PROGRAM main
  VAR
    CONVEYOR_RUN AT %QX0.0 : BOOL;
    PUSHER_EXTEND AT %QX0.1 : BOOL;
    PUSHER_RETRACT AT %QX0.2 : BOOL;
    PASS_LAMP AT %QX0.3 : BOOL;
    FAIL_LAMP AT %QX0.4 : BOOL;
    FAULT_LAMP AT %QX0.5 : BOOL;
    STATION_READY AT %QX0.6 : BOOL;
    SIM_MODE AT %QX2.0 : BOOL := TRUE;
    SIM_UNIT_AT_INSPECTION AT %QX2.1 : BOOL := FALSE;
    SIM_UNIT_AT_REJECT AT %QX2.2 : BOOL := FALSE;
    SIM_VISION_PASS AT %QX2.3 : BOOL := FALSE;
    SIM_VISION_RESULT_VALID AT %QX2.4 : BOOL := FALSE;
    SIM_ESTOP_OK_NC AT %QX2.5 : BOOL := TRUE;
    SIM_GUARD_CLOSED_NC AT %QX2.6 : BOOL := TRUE;
    SIM_AUTO_MODE AT %QX2.7 : BOOL := TRUE;
    SIM_CYCLE_START AT %QX3.0 : BOOL := FALSE;
    SIM_RESET_PB AT %QX3.1 : BOOL := FALSE;
    SIM_PUSHER_EXTENDED AT %QX3.2 : BOOL := FALSE;
    SIM_PUSHER_RETRACTED AT %QX3.3 : BOOL := TRUE;
    SIM_DOWNSTREAM_CLEAR AT %QX3.4 : BOOL := TRUE;
    STATE_CODE AT %QW0 : UINT := 0;
    TOTAL_UNITS AT %QW1 : UINT := 0;
    TOTAL_REJECTS AT %QW2 : UINT := 0;
    LAST_CYCLE_TIME_MS AT %QW3 : UINT := 0;
    FAULT_CODE AT %QW4 : UINT := 0;
    LAST_SERIAL AT %QW5 : UINT := 0;
    LAST_RESULT AT %QW6 : UINT := 0;
    LAST_FAIL_REASON AT %QW7 : UINT := 0;
    SCENARIO_STEP AT %QW8 : UINT := 0;
    SIM_UNIT_SERIAL_IN AT %QW20 : UINT := 0;
    SIM_FAIL_REASON_IN AT %QW21 : UINT := 0;
    S_IDLE : BOOL := TRUE;
    S_READY : BOOL := FALSE;
    S_INSPECTING : BOOL := FALSE;
    S_PASS_RELEASE : BOOL := FALSE;
    S_REJECT_EXTEND : BOOL := FALSE;
    S_REJECT_RETRACT : BOOL := FALSE;
    S_FAULT : BOOL := FALSE;
    IN_UNIT_AT_INSPECTION : BOOL := FALSE;
    IN_UNIT_AT_REJECT : BOOL := FALSE;
    IN_VISION_PASS : BOOL := FALSE;
    IN_VISION_RESULT_VALID : BOOL := FALSE;
    IN_ESTOP_OK_NC : BOOL := FALSE;
    IN_GUARD_CLOSED_NC : BOOL := FALSE;
    IN_AUTO_MODE : BOOL := FALSE;
    IN_CYCLE_START : BOOL := FALSE;
    IN_RESET_PB : BOOL := FALSE;
    IN_PUSHER_EXTENDED : BOOL := FALSE;
    IN_PUSHER_RETRACTED : BOOL := FALSE;
    IN_DOWNSTREAM_CLEAR : BOOL := FALSE;
    START_RISE : BOOL := FALSE;
    START_LAST : BOOL := FALSE;
    RESET_RISE : BOOL := FALSE;
    RESET_LAST : BOOL := FALSE;
    UNIT_RISE : BOOL := FALSE;
    UNIT_LAST : BOOL := FALSE;
    VISION_LAST : BOOL := FALSE;
    VISION_CHANGED : BOOL := FALSE;
    VISION_UNSTABLE_LATCH : BOOL := FALSE;
    RESULT_LATCHED : BOOL := FALSE;
    RESULT_PASS_LATCH : BOOL := FALSE;
    RESULT_FAIL_LATCH : BOOL := FALSE;
    COMPLETE_PULSE : BOOL := FALSE;
    PASS_COMPLETE_PULSE : BOOL := FALSE;
    FAIL_COMPLETE_PULSE : BOOL := FALSE;
    EXTEND_DEMAND : BOOL := FALSE;
    RETRACT_DEMAND : BOOL := FALSE;
    OUTPUT_CONFLICT : BOOL := FALSE;
    FAULT_ESTOP : BOOL := FALSE;
    FAULT_GUARD : BOOL := FALSE;
    FAULT_EXTEND_TIMEOUT : BOOL := FALSE;
    FAULT_RETRACT_TIMEOUT : BOOL := FALSE;
    FAULT_UNIT_STUCK : BOOL := FALSE;
    FAULT_VISION_UNSTABLE : BOOL := FALSE;
    FAULT_OUTPUT_CONFLICT : BOOL := FALSE;
    UNIT_RELEASE_MONITOR : BOOL := FALSE;
    T_VISION_STABLE : TON;
    T_VISION_UNSTABLE : TON;
    T_PASS_RELEASE : TON;
    T_EXTEND_TIMEOUT : TON;
    T_REJECT_SETTLE : TON;
    T_RETRACT_TIMEOUT : TON;
    T_UNIT_STUCK : TON;
    IN_UNIT_SERIAL : UINT := 0;
    IN_FAIL_REASON : UINT := 0;
    CURRENT_SERIAL : UINT := 0;
    CURRENT_FAIL_REASON : UINT := 0;
    CYCLE_START_MS : UDINT := 0;
    NOW_MS : UDINT := 0;
    ALL_SAFE : BOOL := FALSE;
    TON0 : TON;
    TON1 : TON;
    TON2 : TON;
    TON3 : TON;
    TON4 : TON;
    TON5 : TON;
    TON6 : TON;
    TON7 : TON;
    TON8 : TON;
    TON9 : TON;
  END_VAR

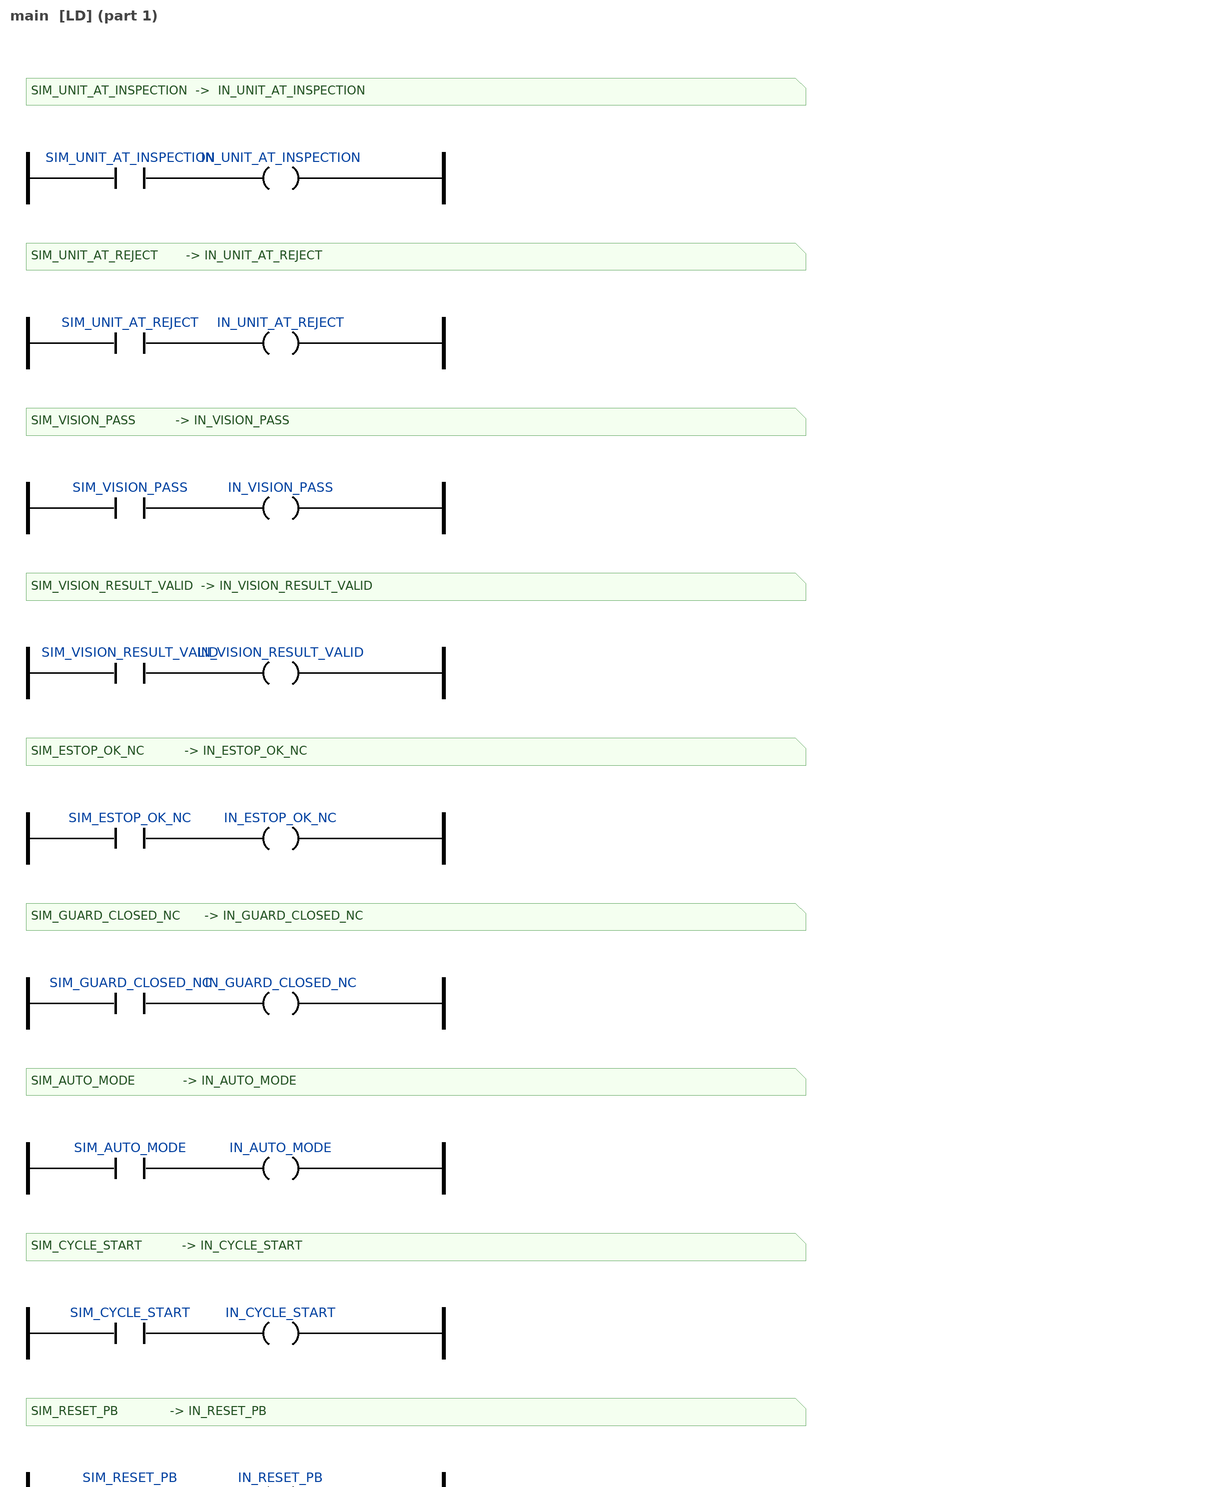
(* LD diagram, written out as Structured Text *)
(* SIM_UNIT_AT_INSPECTION  ->  IN_UNIT_AT_INSPECTION *)
IN_UNIT_AT_INSPECTION := SIM_UNIT_AT_INSPECTION;
(* SIM_UNIT_AT_REJECT       -> IN_UNIT_AT_REJECT *)
IN_UNIT_AT_REJECT := SIM_UNIT_AT_REJECT;
(* SIM_VISION_PASS          -> IN_VISION_PASS *)
IN_VISION_PASS := SIM_VISION_PASS;
(* SIM_VISION_RESULT_VALID  -> IN_VISION_RESULT_VALID *)
IN_VISION_RESULT_VALID := SIM_VISION_RESULT_VALID;
(* SIM_ESTOP_OK_NC          -> IN_ESTOP_OK_NC *)
IN_ESTOP_OK_NC := SIM_ESTOP_OK_NC;
(* SIM_GUARD_CLOSED_NC      -> IN_GUARD_CLOSED_NC *)
IN_GUARD_CLOSED_NC := SIM_GUARD_CLOSED_NC;
(* SIM_AUTO_MODE            -> IN_AUTO_MODE *)
IN_AUTO_MODE := SIM_AUTO_MODE;
(* SIM_CYCLE_START          -> IN_CYCLE_START *)
IN_CYCLE_START := SIM_CYCLE_START;
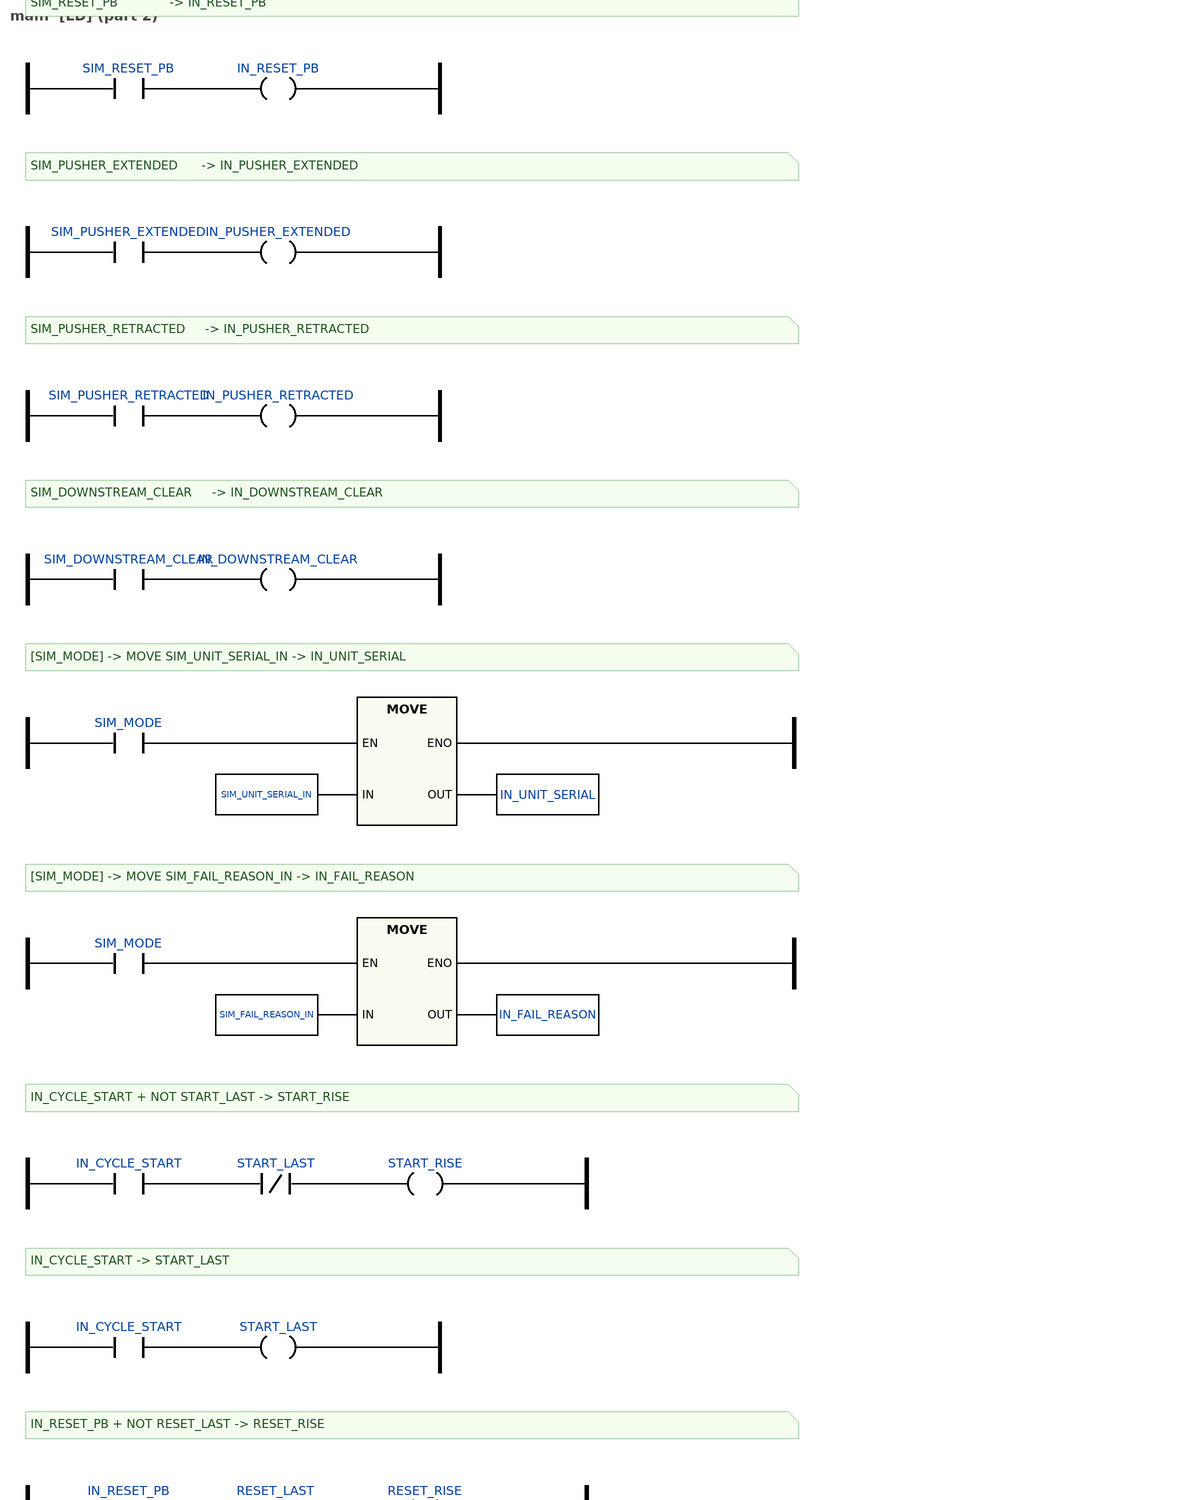
(* SIM_RESET_PB             -> IN_RESET_PB *)
IN_RESET_PB := SIM_RESET_PB;
(* SIM_PUSHER_EXTENDED      -> IN_PUSHER_EXTENDED *)
IN_PUSHER_EXTENDED := SIM_PUSHER_EXTENDED;
(* SIM_PUSHER_RETRACTED     -> IN_PUSHER_RETRACTED *)
IN_PUSHER_RETRACTED := SIM_PUSHER_RETRACTED;
(* SIM_DOWNSTREAM_CLEAR     -> IN_DOWNSTREAM_CLEAR *)
IN_DOWNSTREAM_CLEAR := SIM_DOWNSTREAM_CLEAR;
(* [SIM_MODE] -> MOVE SIM_UNIT_SERIAL_IN -> IN_UNIT_SERIAL *)
IF SIM_MODE THEN IN_UNIT_SERIAL := SIM_UNIT_SERIAL_IN; END_IF;
(* [SIM_MODE] -> MOVE SIM_FAIL_REASON_IN -> IN_FAIL_REASON *)
IF SIM_MODE THEN IN_FAIL_REASON := SIM_FAIL_REASON_IN; END_IF;
(* IN_CYCLE_START + NOT START_LAST -> START_RISE *)
START_RISE := IN_CYCLE_START AND NOT START_LAST;
(* IN_CYCLE_START -> START_LAST *)
START_LAST := IN_CYCLE_START;
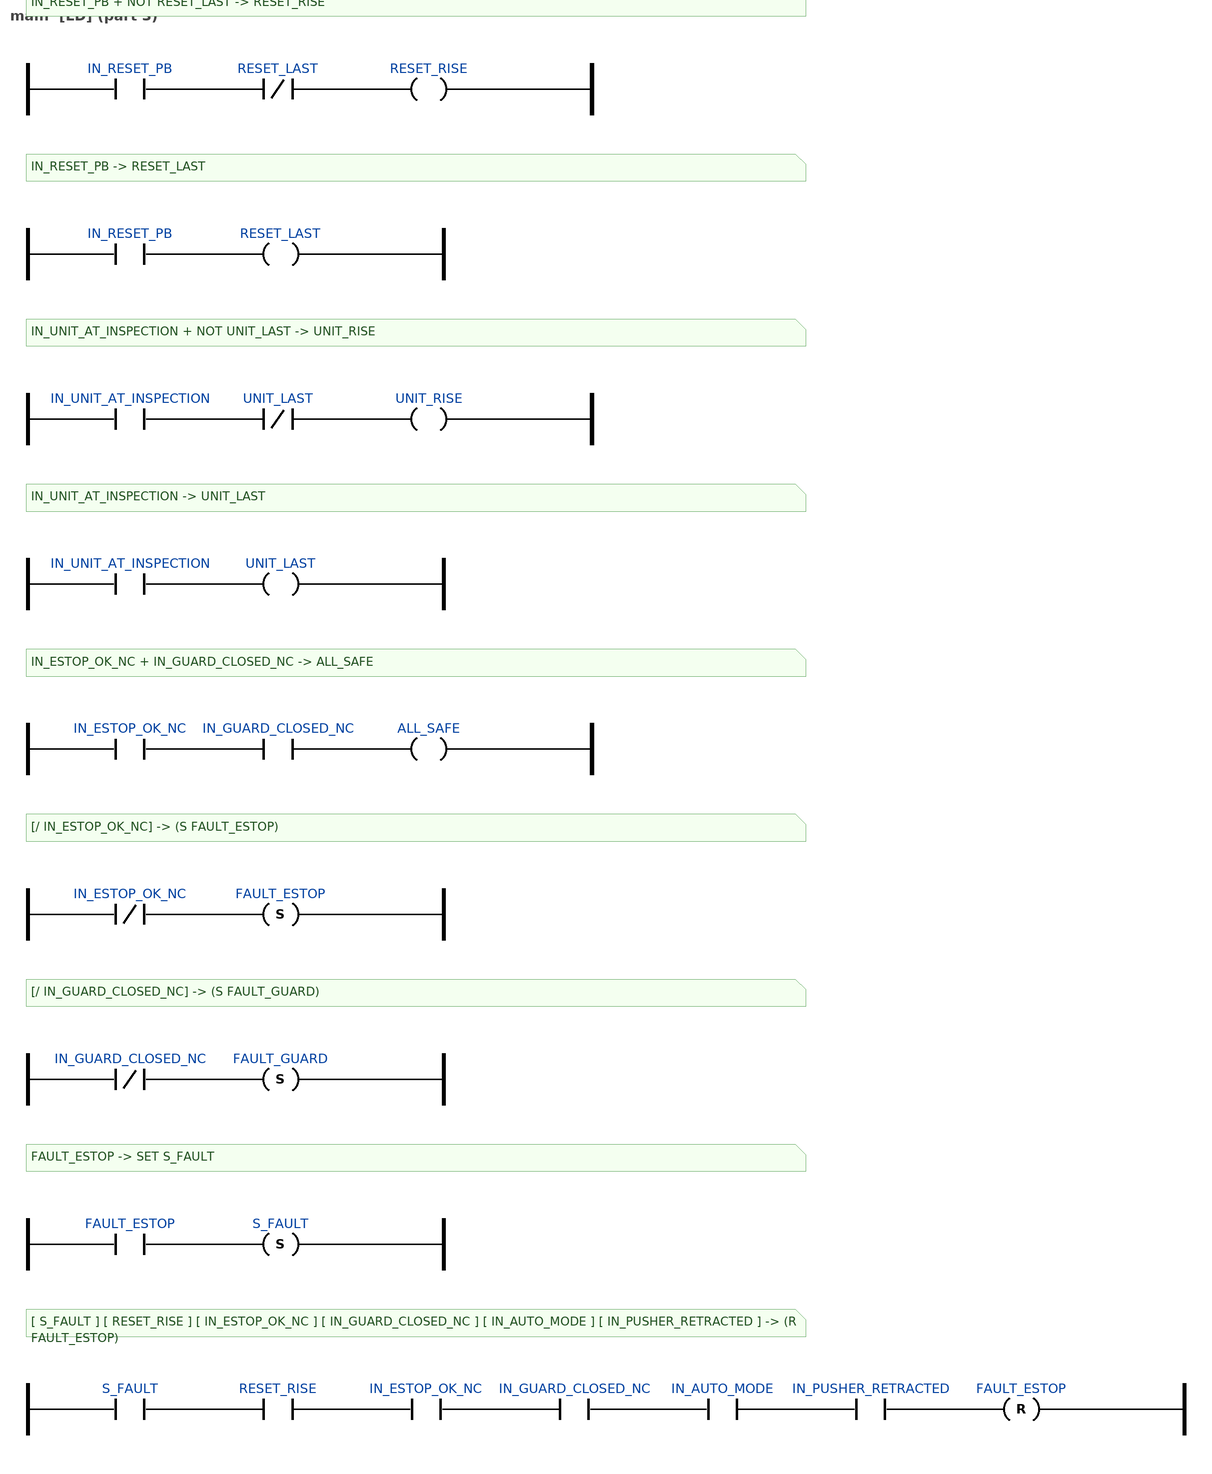
(* IN_RESET_PB + NOT RESET_LAST -> RESET_RISE *)
RESET_RISE := IN_RESET_PB AND NOT RESET_LAST;
(* IN_RESET_PB -> RESET_LAST *)
RESET_LAST := IN_RESET_PB;
(* IN_UNIT_AT_INSPECTION + NOT UNIT_LAST -> UNIT_RISE *)
UNIT_RISE := IN_UNIT_AT_INSPECTION AND NOT UNIT_LAST;
(* IN_UNIT_AT_INSPECTION -> UNIT_LAST *)
UNIT_LAST := IN_UNIT_AT_INSPECTION;
(* IN_ESTOP_OK_NC + IN_GUARD_CLOSED_NC -> ALL_SAFE *)
ALL_SAFE := IN_ESTOP_OK_NC AND IN_GUARD_CLOSED_NC;
(* [/ IN_ESTOP_OK_NC] -> (S FAULT_ESTOP) *)
IF NOT IN_ESTOP_OK_NC THEN FAULT_ESTOP := TRUE; END_IF;
(* [/ IN_GUARD_CLOSED_NC] -> (S FAULT_GUARD) *)
IF NOT IN_GUARD_CLOSED_NC THEN FAULT_GUARD := TRUE; END_IF;
(* FAULT_ESTOP -> SET S_FAULT *)
IF FAULT_ESTOP THEN S_FAULT := TRUE; END_IF;
(* [ S_FAULT ] [ RESET_RISE ] [ IN_ESTOP_OK_NC ] [ IN_GUARD_CLOSED_NC ] [ IN_AUTO_MODE ] [ IN_PUSHER_RETRACTED ] -> (R FAULT_ESTOP) *)
IF S_FAULT AND RESET_RISE AND IN_ESTOP_OK_NC AND IN_GUARD_CLOSED_NC AND IN_AUTO_MODE AND IN_PUSHER_RETRACTED THEN FAULT_ESTOP := FALSE; END_IF;
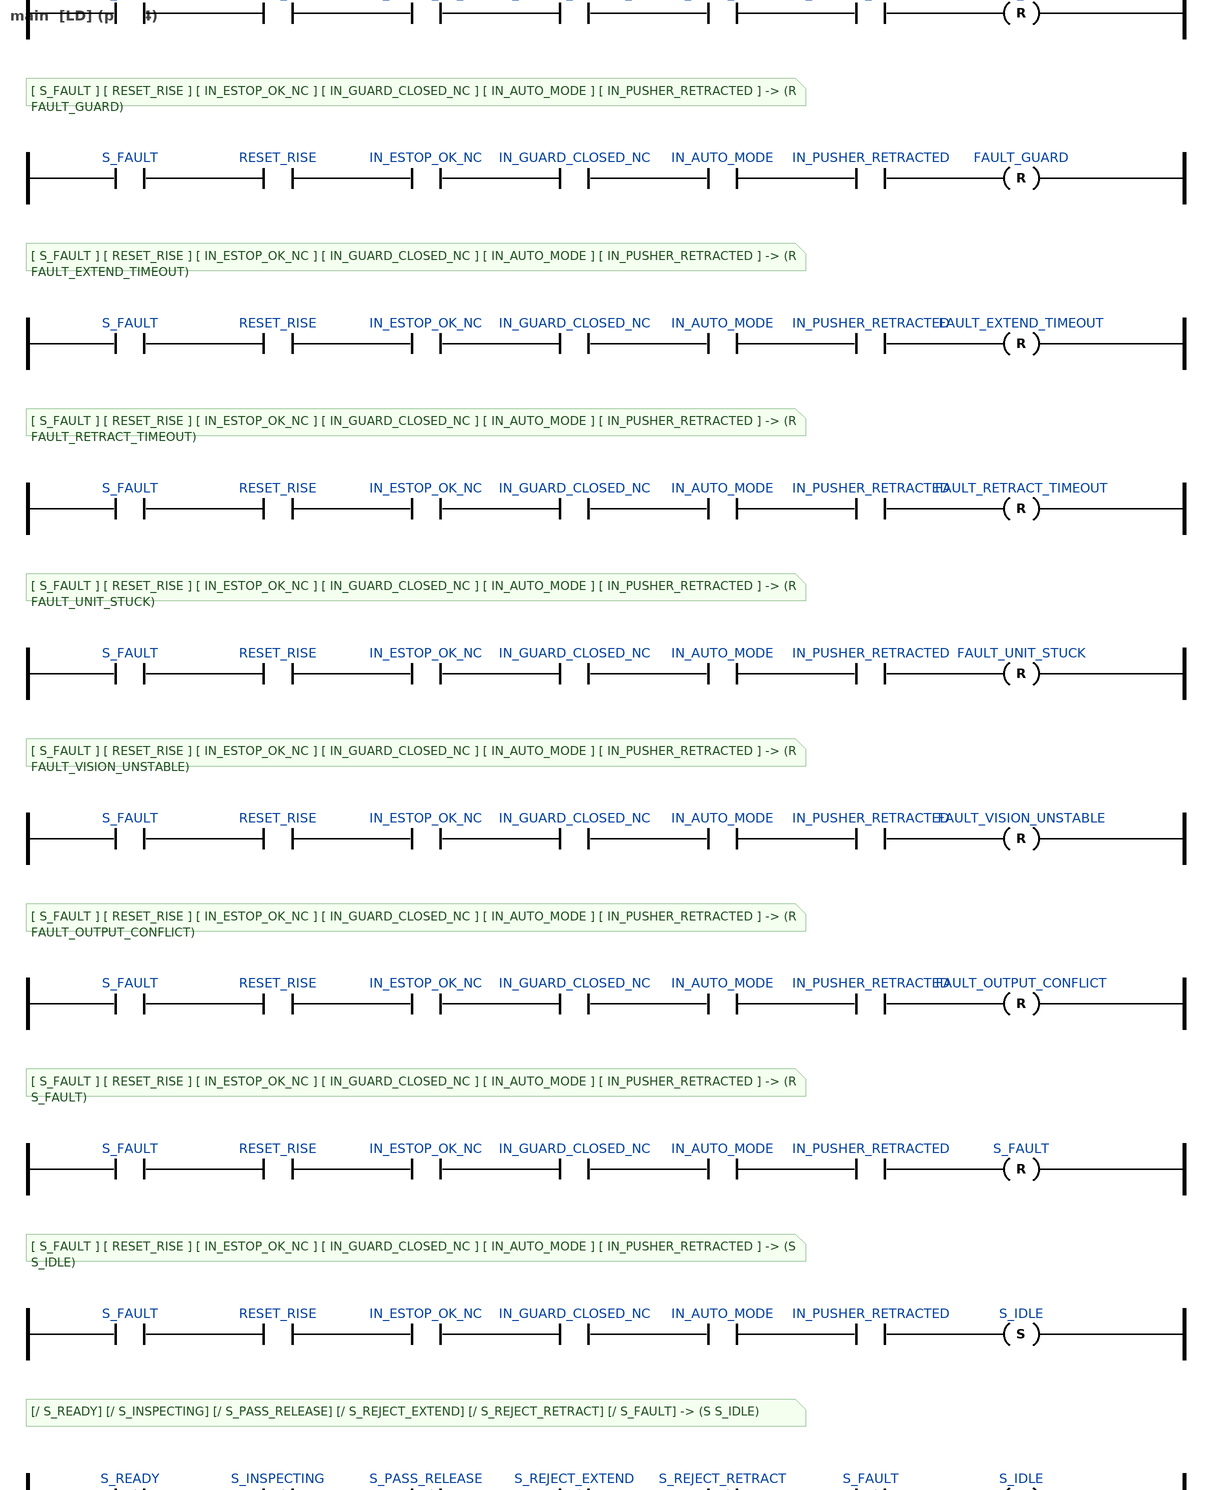
(* [ S_FAULT ] [ RESET_RISE ] [ IN_ESTOP_OK_NC ] [ IN_GUARD_CLOSED_NC ] [ IN_AUTO_MODE ] [ IN_PUSHER_RETRACTED ] -> (R FAULT_GUARD) *)
IF S_FAULT AND RESET_RISE AND IN_ESTOP_OK_NC AND IN_GUARD_CLOSED_NC AND IN_AUTO_MODE AND IN_PUSHER_RETRACTED THEN FAULT_GUARD := FALSE; END_IF;
(* [ S_FAULT ] [ RESET_RISE ] [ IN_ESTOP_OK_NC ] [ IN_GUARD_CLOSED_NC ] [ IN_AUTO_MODE ] [ IN_PUSHER_RETRACTED ] -> (R FAULT_EXTEND_TIMEOUT) *)
IF S_FAULT AND RESET_RISE AND IN_ESTOP_OK_NC AND IN_GUARD_CLOSED_NC AND IN_AUTO_MODE AND IN_PUSHER_RETRACTED THEN FAULT_EXTEND_TIMEOUT := FALSE; END_IF;
(* [ S_FAULT ] [ RESET_RISE ] [ IN_ESTOP_OK_NC ] [ IN_GUARD_CLOSED_NC ] [ IN_AUTO_MODE ] [ IN_PUSHER_RETRACTED ] -> (R FAULT_RETRACT_TIMEOUT) *)
IF S_FAULT AND RESET_RISE AND IN_ESTOP_OK_NC AND IN_GUARD_CLOSED_NC AND IN_AUTO_MODE AND IN_PUSHER_RETRACTED THEN FAULT_RETRACT_TIMEOUT := FALSE; END_IF;
(* [ S_FAULT ] [ RESET_RISE ] [ IN_ESTOP_OK_NC ] [ IN_GUARD_CLOSED_NC ] [ IN_AUTO_MODE ] [ IN_PUSHER_RETRACTED ] -> (R FAULT_UNIT_STUCK) *)
IF S_FAULT AND RESET_RISE AND IN_ESTOP_OK_NC AND IN_GUARD_CLOSED_NC AND IN_AUTO_MODE AND IN_PUSHER_RETRACTED THEN FAULT_UNIT_STUCK := FALSE; END_IF;
(* [ S_FAULT ] [ RESET_RISE ] [ IN_ESTOP_OK_NC ] [ IN_GUARD_CLOSED_NC ] [ IN_AUTO_MODE ] [ IN_PUSHER_RETRACTED ] -> (R FAULT_VISION_UNSTABLE) *)
IF S_FAULT AND RESET_RISE AND IN_ESTOP_OK_NC AND IN_GUARD_CLOSED_NC AND IN_AUTO_MODE AND IN_PUSHER_RETRACTED THEN FAULT_VISION_UNSTABLE := FALSE; END_IF;
(* [ S_FAULT ] [ RESET_RISE ] [ IN_ESTOP_OK_NC ] [ IN_GUARD_CLOSED_NC ] [ IN_AUTO_MODE ] [ IN_PUSHER_RETRACTED ] -> (R FAULT_OUTPUT_CONFLICT) *)
IF S_FAULT AND RESET_RISE AND IN_ESTOP_OK_NC AND IN_GUARD_CLOSED_NC AND IN_AUTO_MODE AND IN_PUSHER_RETRACTED THEN FAULT_OUTPUT_CONFLICT := FALSE; END_IF;
(* [ S_FAULT ] [ RESET_RISE ] [ IN_ESTOP_OK_NC ] [ IN_GUARD_CLOSED_NC ] [ IN_AUTO_MODE ] [ IN_PUSHER_RETRACTED ] -> (R S_FAULT) *)
IF S_FAULT AND RESET_RISE AND IN_ESTOP_OK_NC AND IN_GUARD_CLOSED_NC AND IN_AUTO_MODE AND IN_PUSHER_RETRACTED THEN S_FAULT := FALSE; END_IF;
(* [ S_FAULT ] [ RESET_RISE ] [ IN_ESTOP_OK_NC ] [ IN_GUARD_CLOSED_NC ] [ IN_AUTO_MODE ] [ IN_PUSHER_RETRACTED ] -> (S S_IDLE) *)
IF S_FAULT AND RESET_RISE AND IN_ESTOP_OK_NC AND IN_GUARD_CLOSED_NC AND IN_AUTO_MODE AND IN_PUSHER_RETRACTED THEN S_IDLE := TRUE; END_IF;
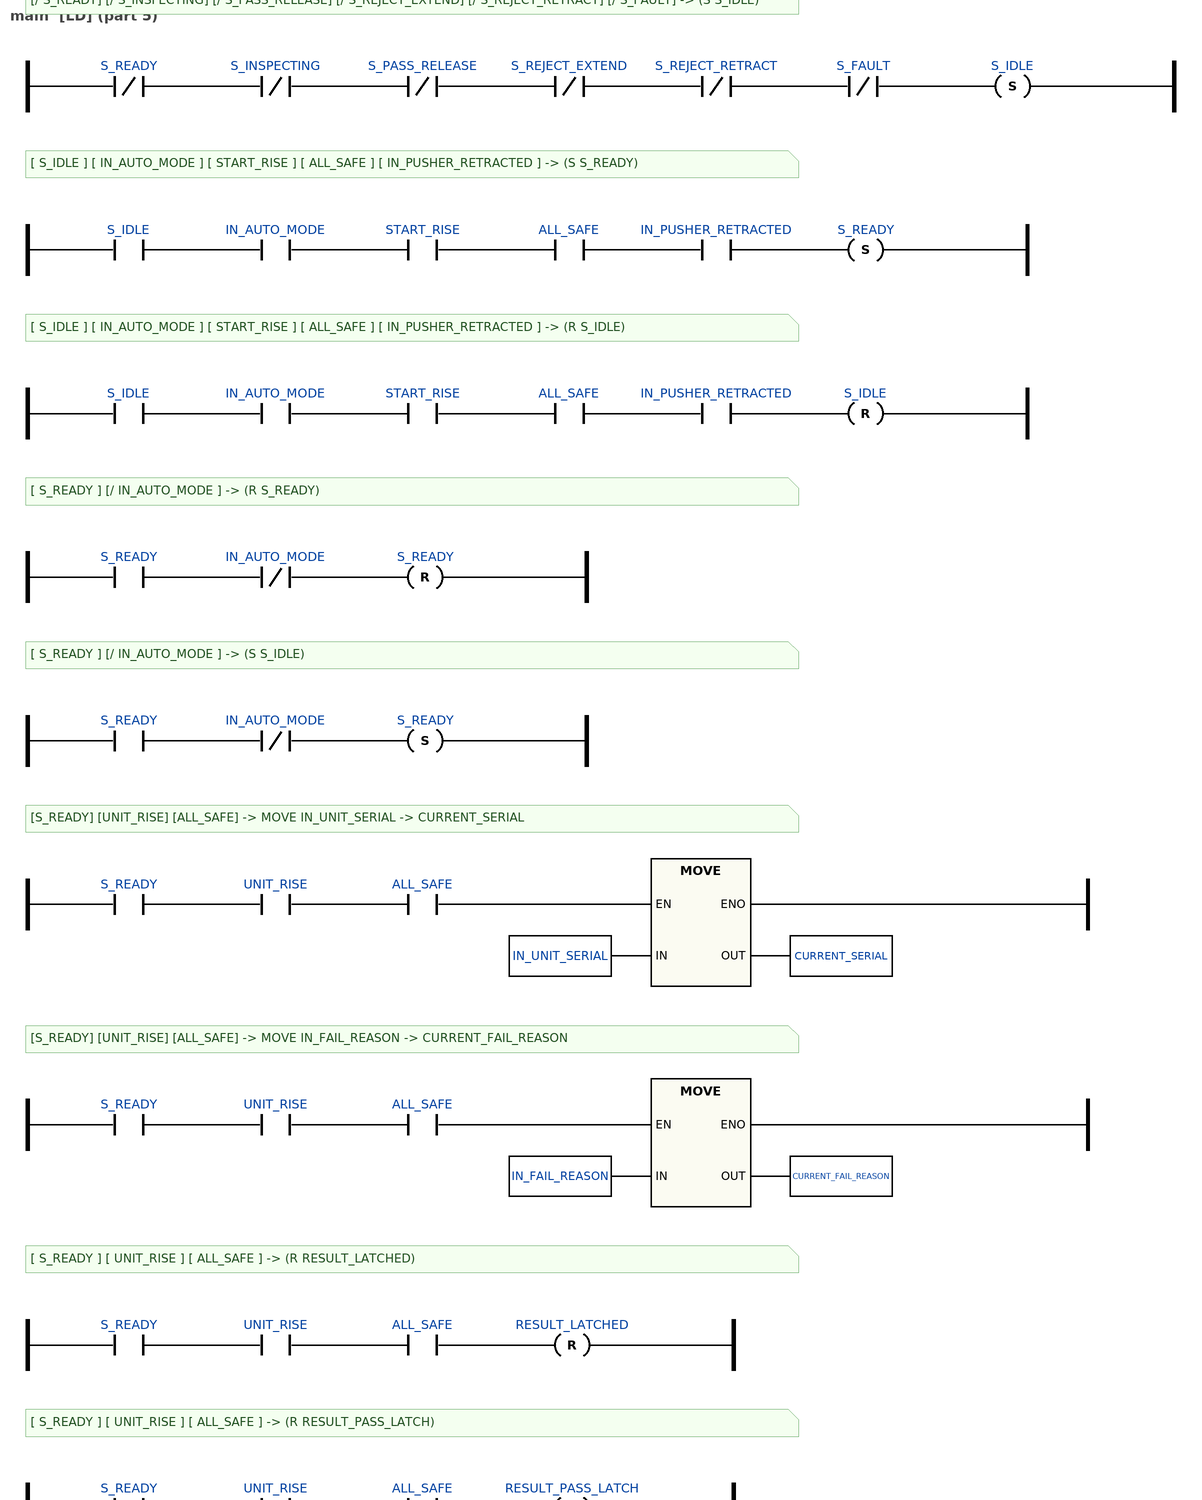
(* [/ S_READY] [/ S_INSPECTING] [/ S_PASS_RELEASE] [/ S_REJECT_EXTEND] [/ S_REJECT_RETRACT] [/ S_FAULT] -> (S S_IDLE) *)
IF NOT S_READY AND NOT S_INSPECTING AND NOT S_PASS_RELEASE AND NOT S_REJECT_EXTEND AND NOT S_REJECT_RETRACT AND NOT S_FAULT THEN S_IDLE := TRUE; END_IF;
(* [ S_IDLE ] [ IN_AUTO_MODE ] [ START_RISE ] [ ALL_SAFE ] [ IN_PUSHER_RETRACTED ] -> (S S_READY) *)
IF S_IDLE AND IN_AUTO_MODE AND START_RISE AND ALL_SAFE AND IN_PUSHER_RETRACTED THEN S_READY := TRUE; END_IF;
(* [ S_IDLE ] [ IN_AUTO_MODE ] [ START_RISE ] [ ALL_SAFE ] [ IN_PUSHER_RETRACTED ] -> (R S_IDLE) *)
IF S_IDLE AND IN_AUTO_MODE AND START_RISE AND ALL_SAFE AND IN_PUSHER_RETRACTED THEN S_IDLE := FALSE; END_IF;
(* [ S_READY ] [/ IN_AUTO_MODE ] -> (R S_READY) *)
IF S_READY AND NOT IN_AUTO_MODE THEN S_READY := FALSE; END_IF;
(* [ S_READY ] [/ IN_AUTO_MODE ] -> (S S_IDLE) *)
IF S_READY AND NOT IN_AUTO_MODE THEN S_READY := TRUE; END_IF;
(* [S_READY] [UNIT_RISE] [ALL_SAFE] -> MOVE IN_UNIT_SERIAL -> CURRENT_SERIAL *)
IF S_READY AND UNIT_RISE AND ALL_SAFE THEN CURRENT_SERIAL := IN_UNIT_SERIAL; END_IF;
(* [S_READY] [UNIT_RISE] [ALL_SAFE] -> MOVE IN_FAIL_REASON -> CURRENT_FAIL_REASON *)
IF S_READY AND UNIT_RISE AND ALL_SAFE THEN CURRENT_FAIL_REASON := IN_FAIL_REASON; END_IF;
(* [ S_READY ] [ UNIT_RISE ] [ ALL_SAFE ] -> (R RESULT_LATCHED) *)
IF S_READY AND UNIT_RISE AND ALL_SAFE THEN RESULT_LATCHED := FALSE; END_IF;
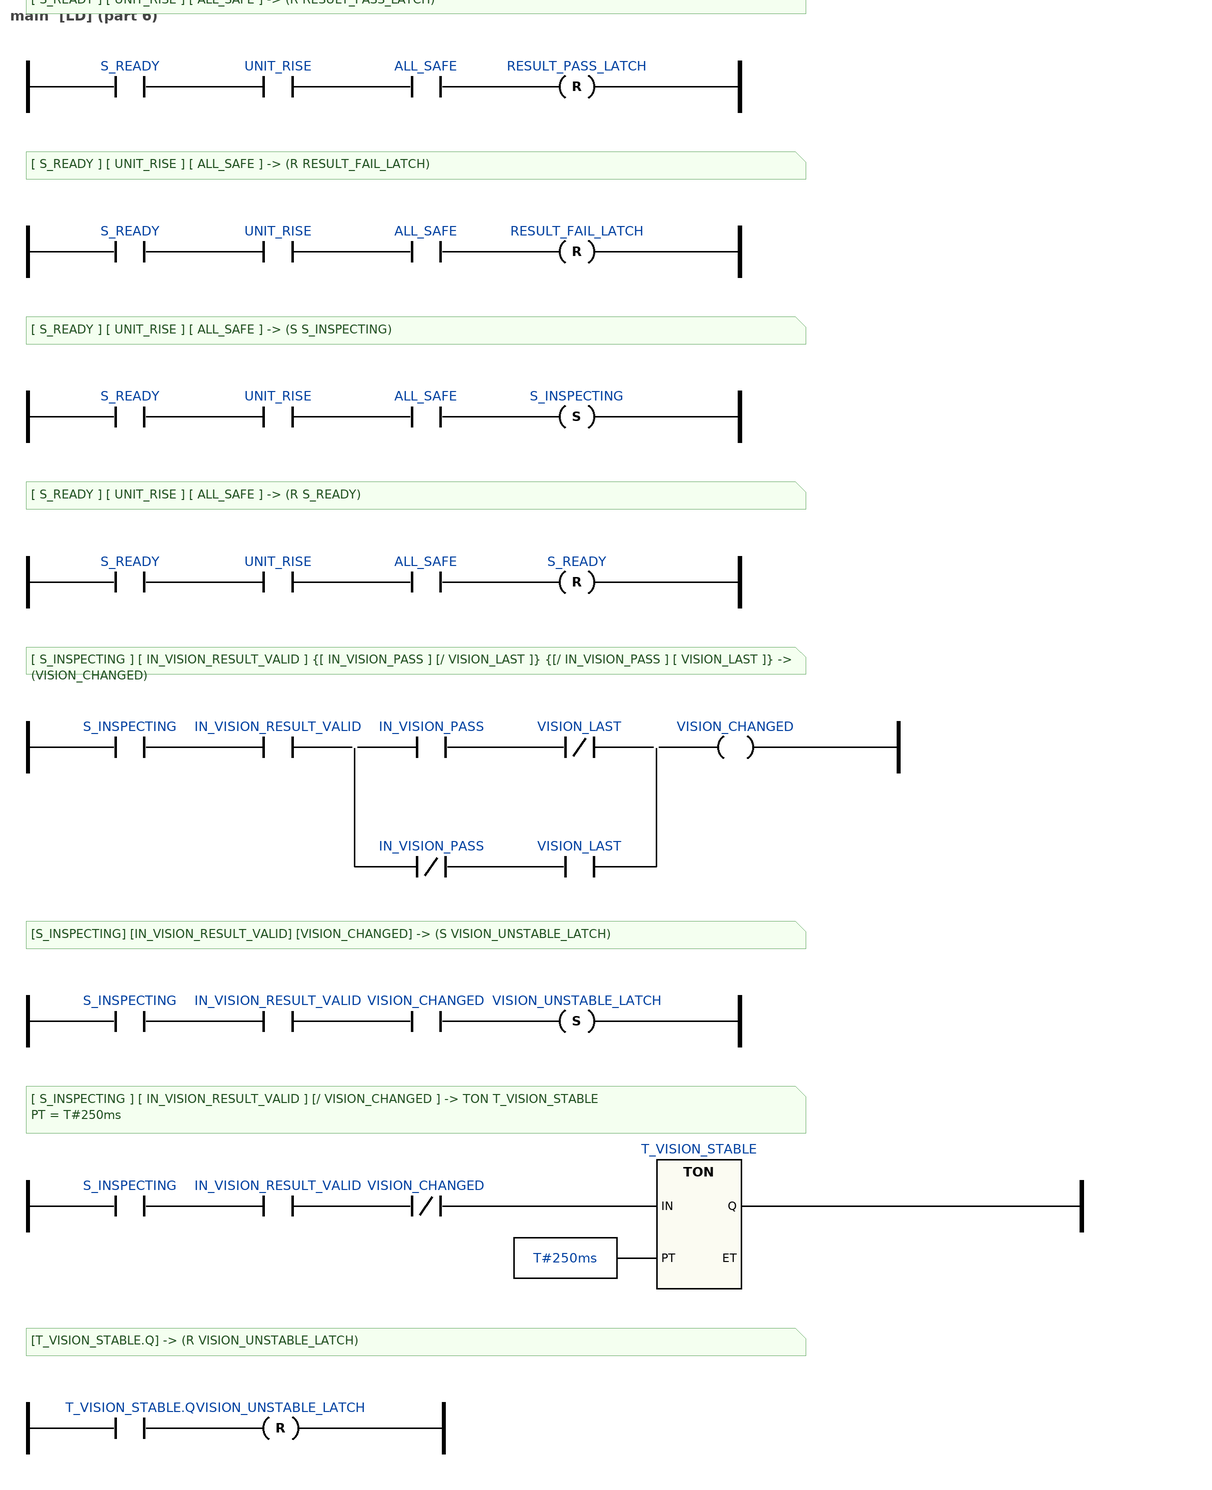
(* [ S_READY ] [ UNIT_RISE ] [ ALL_SAFE ] -> (R RESULT_PASS_LATCH) *)
IF S_READY AND UNIT_RISE AND ALL_SAFE THEN RESULT_PASS_LATCH := FALSE; END_IF;
(* [ S_READY ] [ UNIT_RISE ] [ ALL_SAFE ] -> (R RESULT_FAIL_LATCH) *)
IF S_READY AND UNIT_RISE AND ALL_SAFE THEN RESULT_FAIL_LATCH := FALSE; END_IF;
(* [ S_READY ] [ UNIT_RISE ] [ ALL_SAFE ] -> (S S_INSPECTING) *)
IF S_READY AND UNIT_RISE AND ALL_SAFE THEN S_INSPECTING := TRUE; END_IF;
(* [ S_READY ] [ UNIT_RISE ] [ ALL_SAFE ] -> (R S_READY) *)
IF S_READY AND UNIT_RISE AND ALL_SAFE THEN S_READY := FALSE; END_IF;
(* [ S_INSPECTING ] [ IN_VISION_RESULT_VALID ] {[ IN_VISION_PASS ] [/ VISION_LAST ]} {[/ IN_VISION_PASS ] [ VISION_LAST ]} -> (VISION_CHANGED) *)
VISION_CHANGED := S_INSPECTING AND IN_VISION_RESULT_VALID AND (NOT IN_VISION_PASS AND VISION_LAST OR IN_VISION_PASS AND NOT VISION_LAST);
(* [S_INSPECTING] [IN_VISION_RESULT_VALID] [VISION_CHANGED] -> (S VISION_UNSTABLE_LATCH) *)
IF S_INSPECTING AND IN_VISION_RESULT_VALID AND VISION_CHANGED THEN VISION_UNSTABLE_LATCH := TRUE; END_IF;
(* [ S_INSPECTING ] [ IN_VISION_RESULT_VALID ] [/ VISION_CHANGED ] -> TON T_VISION_STABLE
PT = T#250ms *)
(* [T_VISION_STABLE.Q] -> (R VISION_UNSTABLE_LATCH) *)
IF T_VISION_STABLE.Q THEN VISION_UNSTABLE_LATCH := FALSE; END_IF;
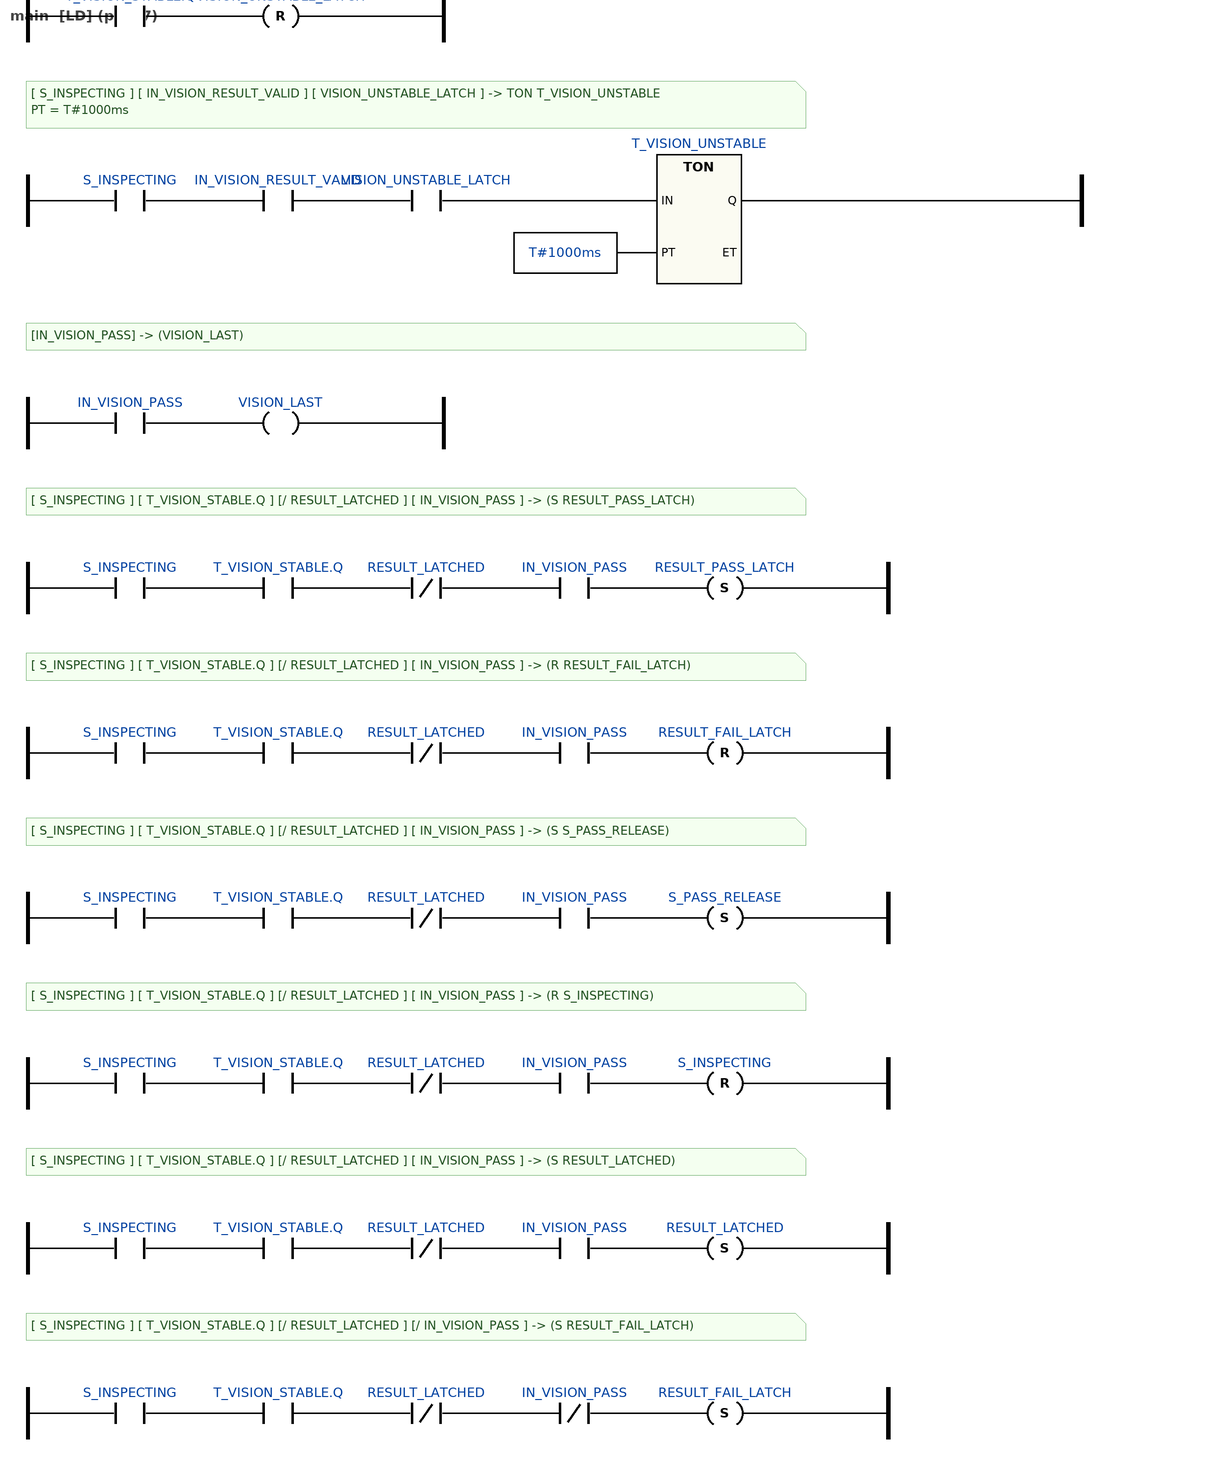
(* [ S_INSPECTING ] [ IN_VISION_RESULT_VALID ] [ VISION_UNSTABLE_LATCH ] -> TON T_VISION_UNSTABLE
PT = T#1000ms *)
(* [IN_VISION_PASS] -> (VISION_LAST) *)
VISION_LAST := IN_VISION_PASS;
(* [ S_INSPECTING ] [ T_VISION_STABLE.Q ] [/ RESULT_LATCHED ] [ IN_VISION_PASS ] -> (S RESULT_PASS_LATCH) *)
IF S_INSPECTING AND T_VISION_STABLE.Q AND NOT RESULT_LATCHED AND IN_VISION_PASS THEN RESULT_PASS_LATCH := TRUE; END_IF;
(* [ S_INSPECTING ] [ T_VISION_STABLE.Q ] [/ RESULT_LATCHED ] [ IN_VISION_PASS ] -> (R RESULT_FAIL_LATCH) *)
IF S_INSPECTING AND T_VISION_STABLE.Q AND NOT RESULT_LATCHED AND IN_VISION_PASS THEN RESULT_FAIL_LATCH := FALSE; END_IF;
(* [ S_INSPECTING ] [ T_VISION_STABLE.Q ] [/ RESULT_LATCHED ] [ IN_VISION_PASS ] -> (S S_PASS_RELEASE) *)
IF S_INSPECTING AND T_VISION_STABLE.Q AND NOT RESULT_LATCHED AND IN_VISION_PASS THEN S_PASS_RELEASE := TRUE; END_IF;
(* [ S_INSPECTING ] [ T_VISION_STABLE.Q ] [/ RESULT_LATCHED ] [ IN_VISION_PASS ] -> (R S_INSPECTING) *)
IF S_INSPECTING AND T_VISION_STABLE.Q AND NOT RESULT_LATCHED AND IN_VISION_PASS THEN S_INSPECTING := FALSE; END_IF;
(* [ S_INSPECTING ] [ T_VISION_STABLE.Q ] [/ RESULT_LATCHED ] [ IN_VISION_PASS ] -> (S RESULT_LATCHED) *)
IF S_INSPECTING AND T_VISION_STABLE.Q AND NOT RESULT_LATCHED AND IN_VISION_PASS THEN RESULT_LATCHED := TRUE; END_IF;
(* [ S_INSPECTING ] [ T_VISION_STABLE.Q ] [/ RESULT_LATCHED ] [/ IN_VISION_PASS ] -> (S RESULT_FAIL_LATCH) *)
IF S_INSPECTING AND T_VISION_STABLE.Q AND NOT RESULT_LATCHED AND NOT IN_VISION_PASS THEN RESULT_FAIL_LATCH := TRUE; END_IF;
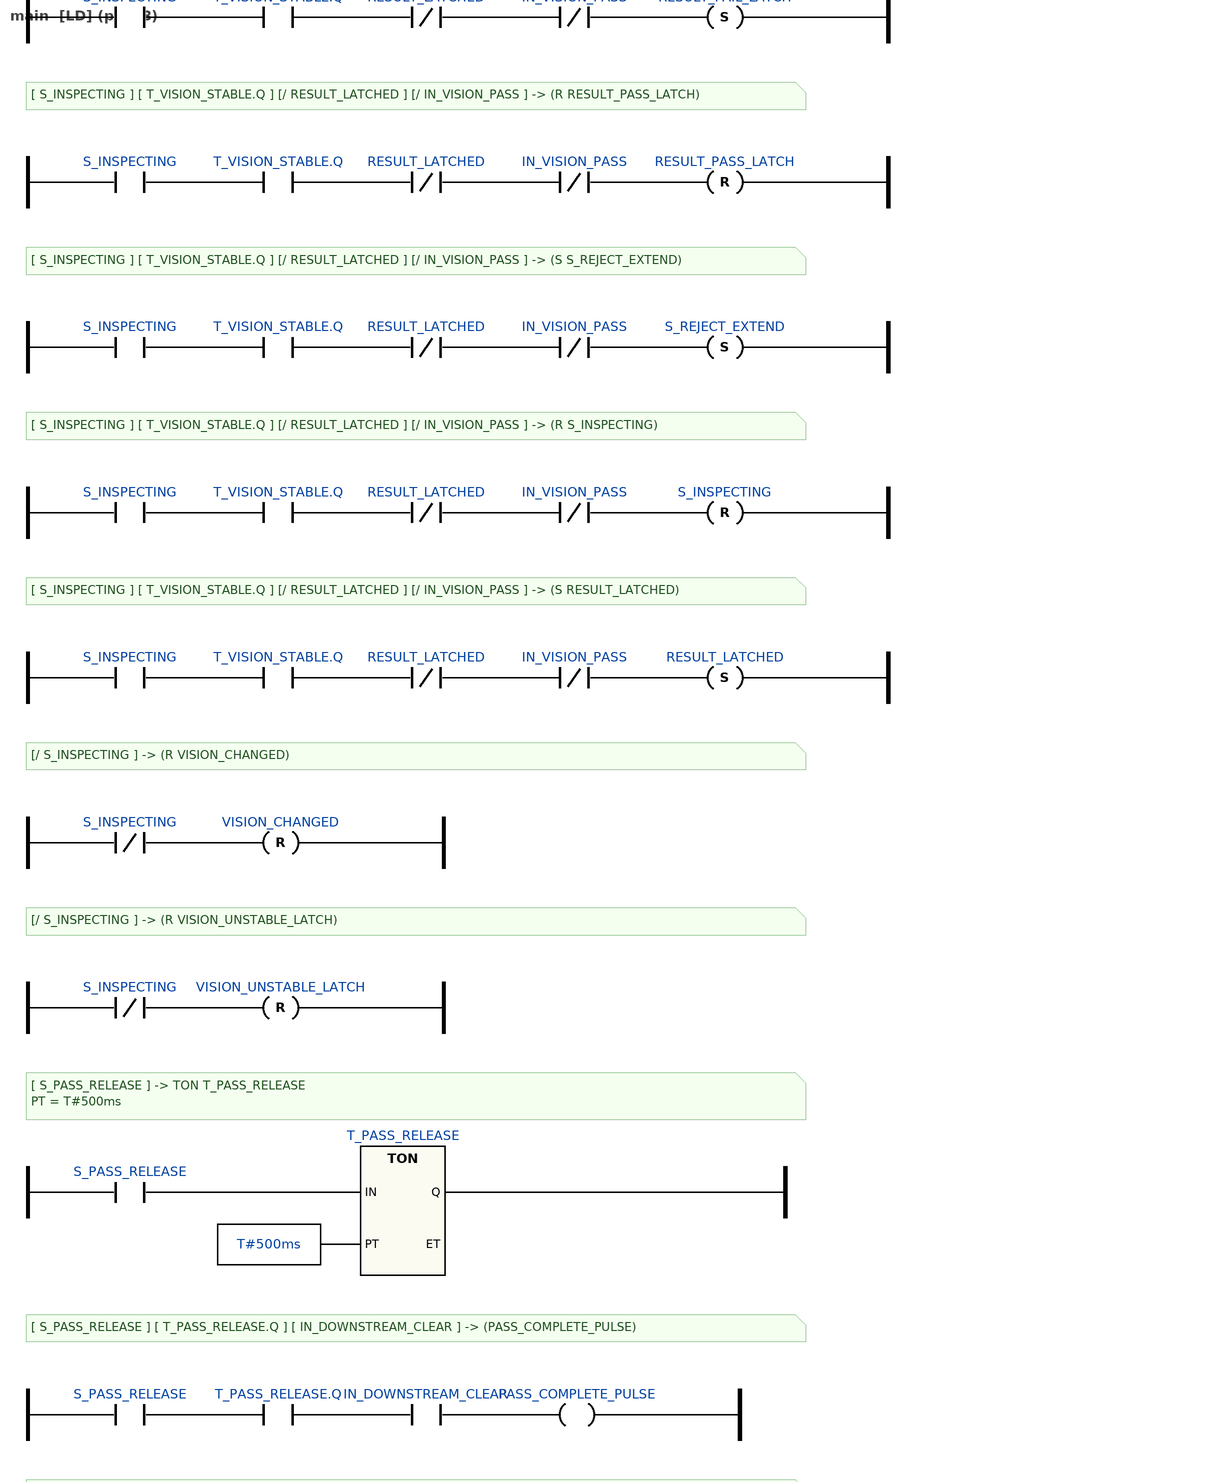
(* [ S_INSPECTING ] [ T_VISION_STABLE.Q ] [/ RESULT_LATCHED ] [/ IN_VISION_PASS ] -> (R RESULT_PASS_LATCH) *)
IF S_INSPECTING AND T_VISION_STABLE.Q AND NOT RESULT_LATCHED AND NOT IN_VISION_PASS THEN RESULT_PASS_LATCH := FALSE; END_IF;
(* [ S_INSPECTING ] [ T_VISION_STABLE.Q ] [/ RESULT_LATCHED ] [/ IN_VISION_PASS ] -> (S S_REJECT_EXTEND) *)
IF S_INSPECTING AND T_VISION_STABLE.Q AND NOT RESULT_LATCHED AND NOT IN_VISION_PASS THEN S_REJECT_EXTEND := TRUE; END_IF;
(* [ S_INSPECTING ] [ T_VISION_STABLE.Q ] [/ RESULT_LATCHED ] [/ IN_VISION_PASS ] -> (R S_INSPECTING) *)
IF S_INSPECTING AND T_VISION_STABLE.Q AND NOT RESULT_LATCHED AND NOT IN_VISION_PASS THEN S_INSPECTING := FALSE; END_IF;
(* [ S_INSPECTING ] [ T_VISION_STABLE.Q ] [/ RESULT_LATCHED ] [/ IN_VISION_PASS ] -> (S RESULT_LATCHED) *)
IF S_INSPECTING AND T_VISION_STABLE.Q AND NOT RESULT_LATCHED AND NOT IN_VISION_PASS THEN RESULT_LATCHED := TRUE; END_IF;
(* [/ S_INSPECTING ] -> (R VISION_CHANGED) *)
IF NOT S_INSPECTING THEN VISION_CHANGED := FALSE; END_IF;
(* [/ S_INSPECTING ] -> (R VISION_UNSTABLE_LATCH) *)
IF NOT S_INSPECTING THEN VISION_UNSTABLE_LATCH := FALSE; END_IF;
(* [ S_PASS_RELEASE ] -> TON T_PASS_RELEASE
PT = T#500ms *)
(* [ S_PASS_RELEASE ] [ T_PASS_RELEASE.Q ] [ IN_DOWNSTREAM_CLEAR ] -> (PASS_COMPLETE_PULSE) *)
PASS_COMPLETE_PULSE := S_PASS_RELEASE AND T_PASS_RELEASE.Q AND IN_DOWNSTREAM_CLEAR;
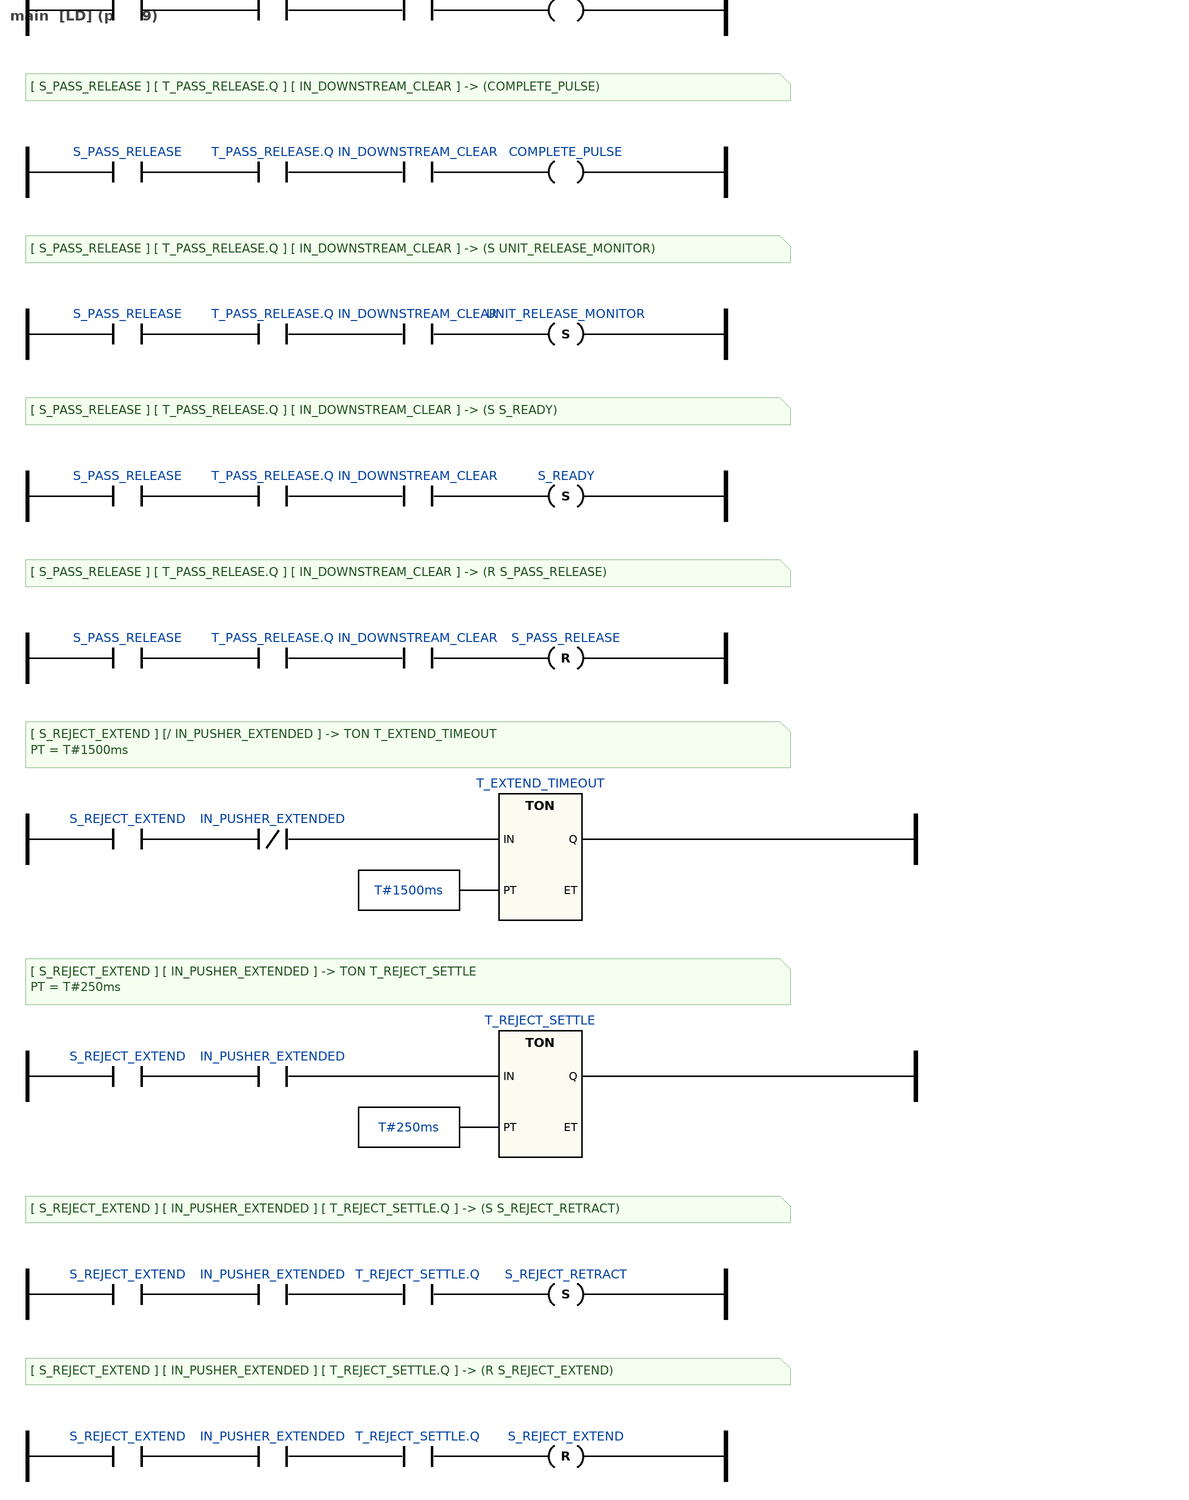
(* [ S_PASS_RELEASE ] [ T_PASS_RELEASE.Q ] [ IN_DOWNSTREAM_CLEAR ] -> (COMPLETE_PULSE) *)
COMPLETE_PULSE := S_PASS_RELEASE AND T_PASS_RELEASE.Q AND IN_DOWNSTREAM_CLEAR;
(* [ S_PASS_RELEASE ] [ T_PASS_RELEASE.Q ] [ IN_DOWNSTREAM_CLEAR ] -> (S UNIT_RELEASE_MONITOR) *)
IF S_PASS_RELEASE AND T_PASS_RELEASE.Q AND IN_DOWNSTREAM_CLEAR THEN UNIT_RELEASE_MONITOR := TRUE; END_IF;
(* [ S_PASS_RELEASE ] [ T_PASS_RELEASE.Q ] [ IN_DOWNSTREAM_CLEAR ] -> (S S_READY) *)
IF S_PASS_RELEASE AND T_PASS_RELEASE.Q AND IN_DOWNSTREAM_CLEAR THEN S_READY := TRUE; END_IF;
(* [ S_PASS_RELEASE ] [ T_PASS_RELEASE.Q ] [ IN_DOWNSTREAM_CLEAR ] -> (R S_PASS_RELEASE) *)
IF S_PASS_RELEASE AND T_PASS_RELEASE.Q AND IN_DOWNSTREAM_CLEAR THEN S_PASS_RELEASE := FALSE; END_IF;
(* [ S_REJECT_EXTEND ] [/ IN_PUSHER_EXTENDED ] -> TON T_EXTEND_TIMEOUT
PT = T#1500ms *)
(* [ S_REJECT_EXTEND ] [ IN_PUSHER_EXTENDED ] -> TON T_REJECT_SETTLE
PT = T#250ms *)
(* [ S_REJECT_EXTEND ] [ IN_PUSHER_EXTENDED ] [ T_REJECT_SETTLE.Q ] -> (S S_REJECT_RETRACT) *)
IF S_REJECT_EXTEND AND IN_PUSHER_EXTENDED AND T_REJECT_SETTLE.Q THEN S_REJECT_RETRACT := TRUE; END_IF;
(* [ S_REJECT_EXTEND ] [ IN_PUSHER_EXTENDED ] [ T_REJECT_SETTLE.Q ] -> (R S_REJECT_EXTEND) *)
IF S_REJECT_EXTEND AND IN_PUSHER_EXTENDED AND T_REJECT_SETTLE.Q THEN S_REJECT_EXTEND := FALSE; END_IF;
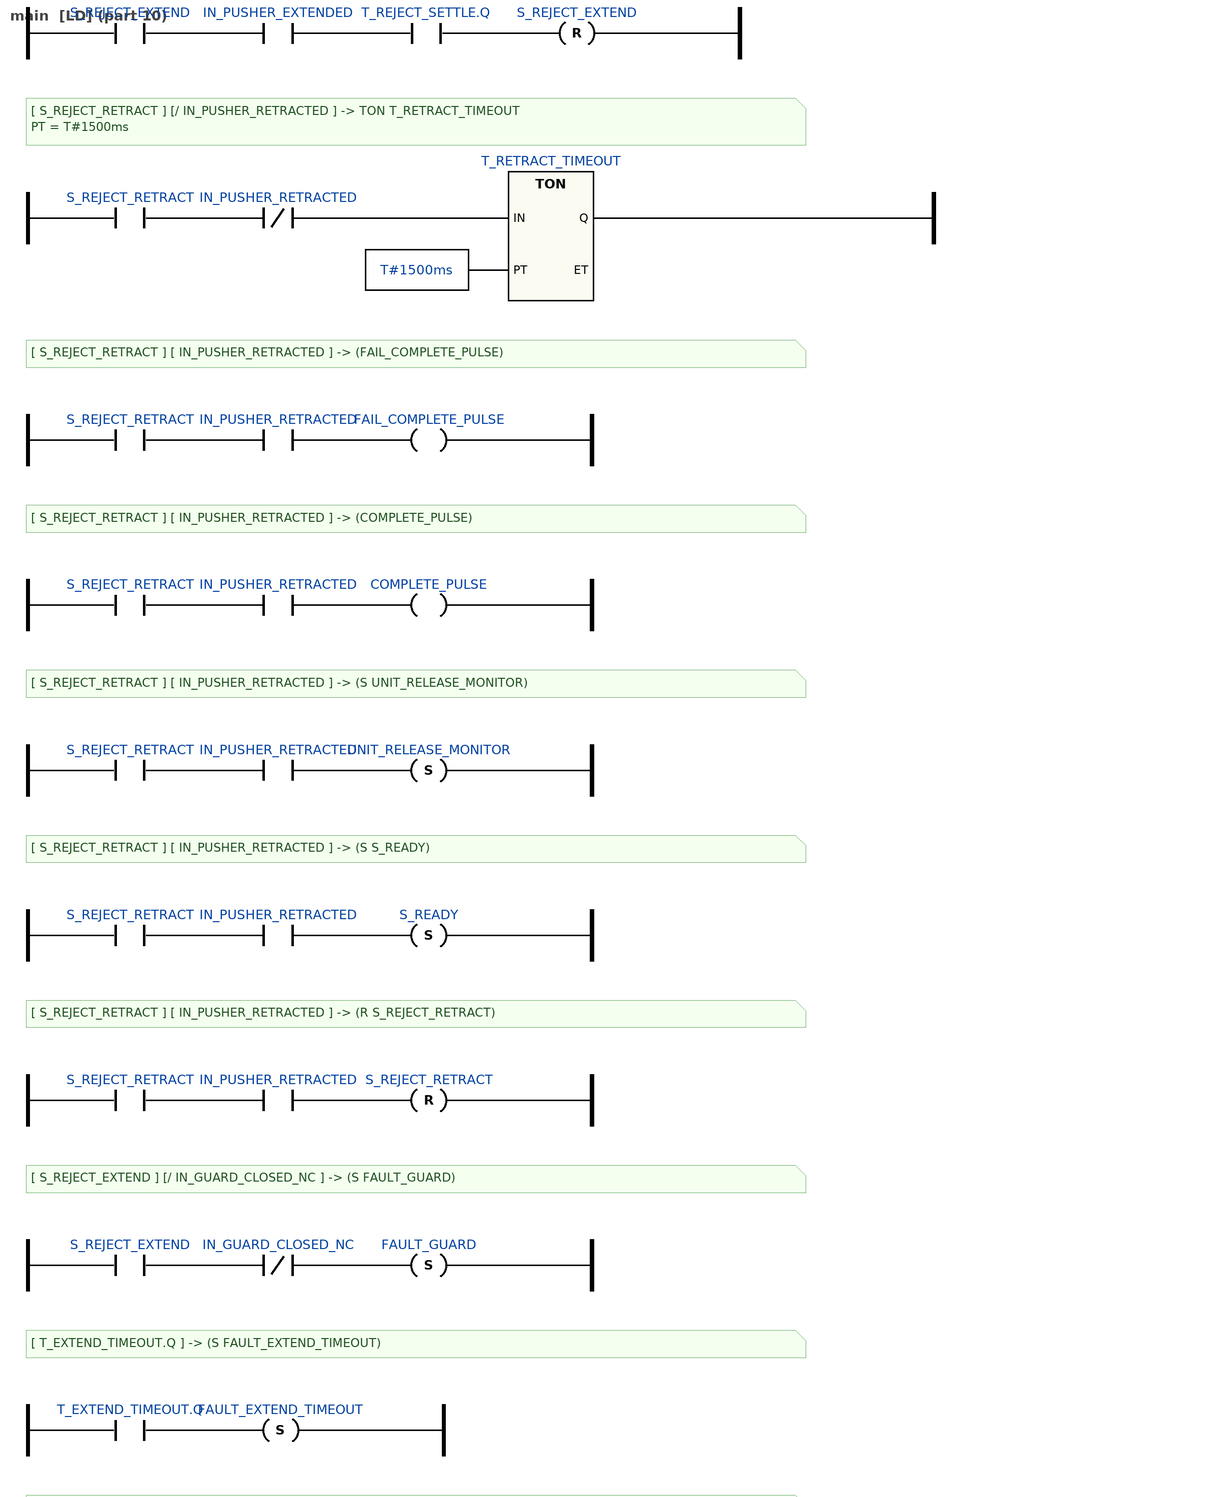
(* [ S_REJECT_RETRACT ] [/ IN_PUSHER_RETRACTED ] -> TON T_RETRACT_TIMEOUT
PT = T#1500ms *)
(* [ S_REJECT_RETRACT ] [ IN_PUSHER_RETRACTED ] -> (FAIL_COMPLETE_PULSE) *)
FAIL_COMPLETE_PULSE := S_REJECT_RETRACT AND IN_PUSHER_RETRACTED;
(* [ S_REJECT_RETRACT ] [ IN_PUSHER_RETRACTED ] -> (COMPLETE_PULSE) *)
COMPLETE_PULSE := S_REJECT_RETRACT AND IN_PUSHER_RETRACTED;
(* [ S_REJECT_RETRACT ] [ IN_PUSHER_RETRACTED ] -> (S UNIT_RELEASE_MONITOR) *)
IF S_REJECT_RETRACT AND IN_PUSHER_RETRACTED THEN UNIT_RELEASE_MONITOR := TRUE; END_IF;
(* [ S_REJECT_RETRACT ] [ IN_PUSHER_RETRACTED ] -> (S S_READY) *)
IF S_REJECT_RETRACT AND IN_PUSHER_RETRACTED THEN S_READY := TRUE; END_IF;
(* [ S_REJECT_RETRACT ] [ IN_PUSHER_RETRACTED ] -> (R S_REJECT_RETRACT) *)
IF S_REJECT_RETRACT AND IN_PUSHER_RETRACTED THEN S_REJECT_RETRACT := FALSE; END_IF;
(* [ S_REJECT_EXTEND ] [/ IN_GUARD_CLOSED_NC ] -> (S FAULT_GUARD) *)
IF S_REJECT_EXTEND AND NOT IN_GUARD_CLOSED_NC THEN FAULT_GUARD := TRUE; END_IF;
(* [ T_EXTEND_TIMEOUT.Q ] -> (S FAULT_EXTEND_TIMEOUT) *)
IF T_EXTEND_TIMEOUT.Q THEN FAULT_EXTEND_TIMEOUT := TRUE; END_IF;
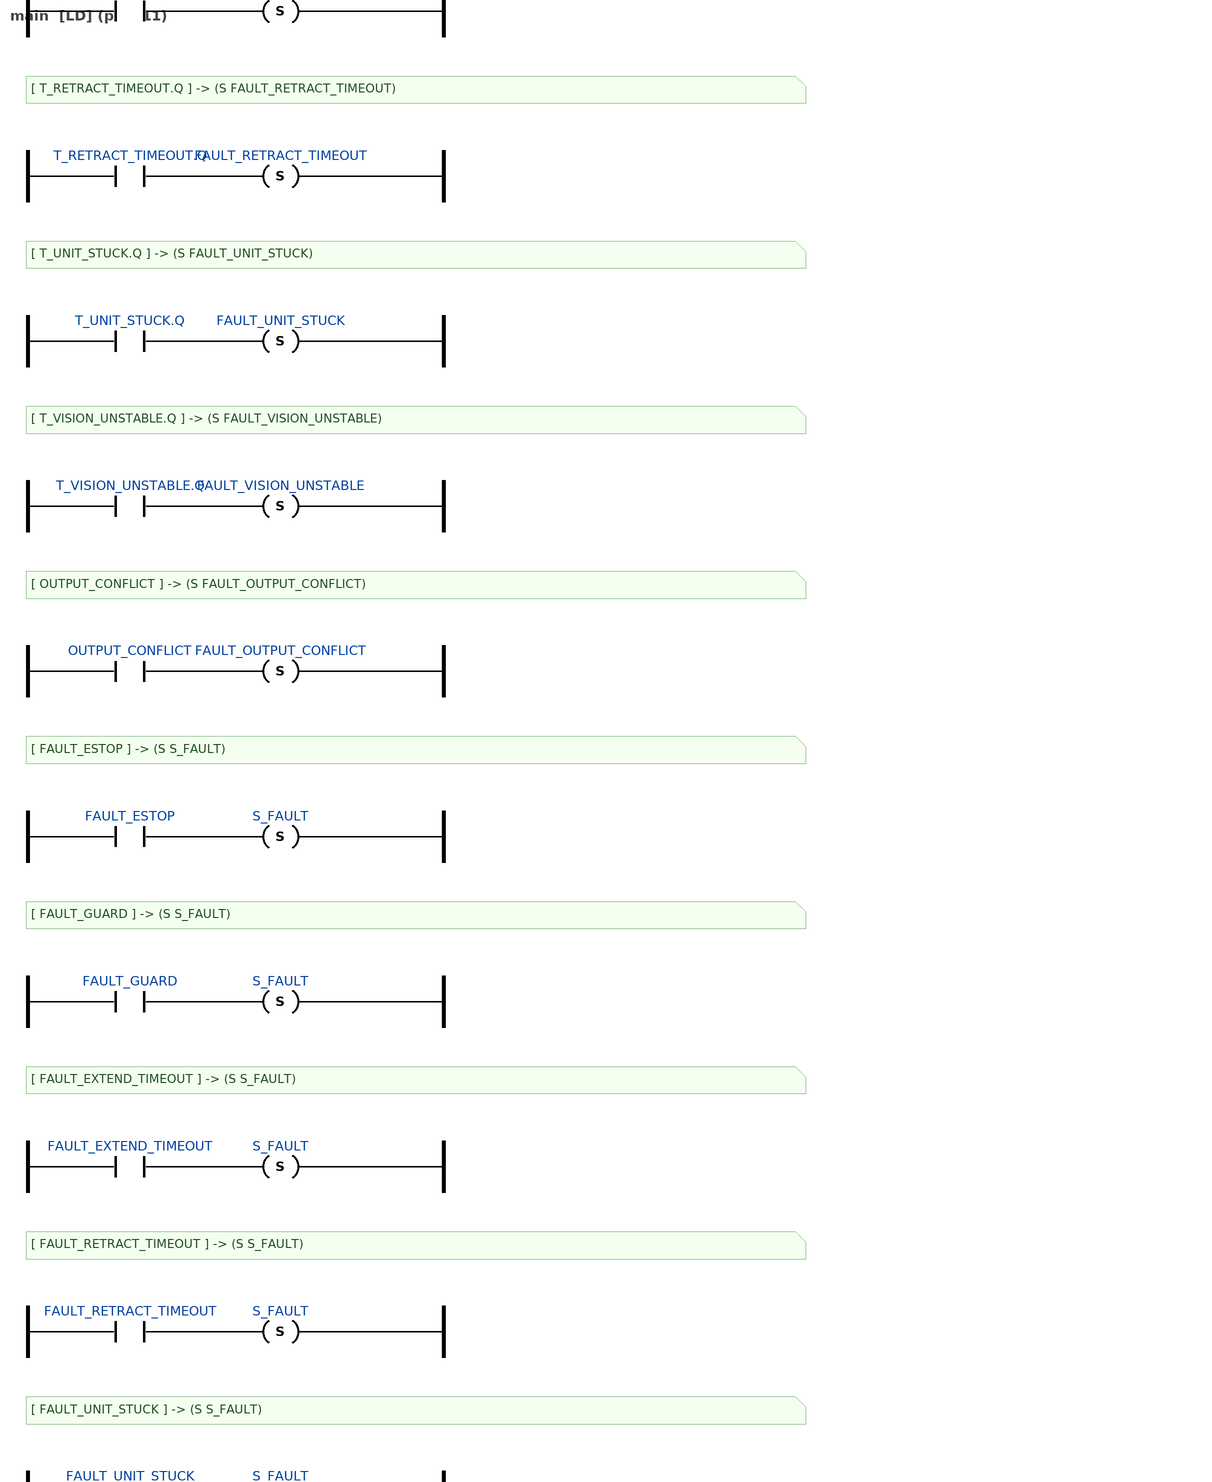
(* [ T_RETRACT_TIMEOUT.Q ] -> (S FAULT_RETRACT_TIMEOUT) *)
IF T_RETRACT_TIMEOUT.Q THEN FAULT_RETRACT_TIMEOUT := TRUE; END_IF;
(* [ T_UNIT_STUCK.Q ] -> (S FAULT_UNIT_STUCK) *)
IF T_UNIT_STUCK.Q THEN FAULT_UNIT_STUCK := TRUE; END_IF;
(* [ T_VISION_UNSTABLE.Q ] -> (S FAULT_VISION_UNSTABLE) *)
IF T_VISION_UNSTABLE.Q THEN FAULT_VISION_UNSTABLE := TRUE; END_IF;
(* [ OUTPUT_CONFLICT ] -> (S FAULT_OUTPUT_CONFLICT) *)
IF OUTPUT_CONFLICT THEN FAULT_OUTPUT_CONFLICT := TRUE; END_IF;
(* [ FAULT_ESTOP ] -> (S S_FAULT) *)
IF FAULT_ESTOP THEN S_FAULT := TRUE; END_IF;
(* [ FAULT_GUARD ] -> (S S_FAULT) *)
IF FAULT_GUARD THEN S_FAULT := TRUE; END_IF;
(* [ FAULT_EXTEND_TIMEOUT ] -> (S S_FAULT) *)
IF FAULT_EXTEND_TIMEOUT THEN S_FAULT := TRUE; END_IF;
(* [ FAULT_RETRACT_TIMEOUT ] -> (S S_FAULT) *)
IF FAULT_RETRACT_TIMEOUT THEN S_FAULT := TRUE; END_IF;
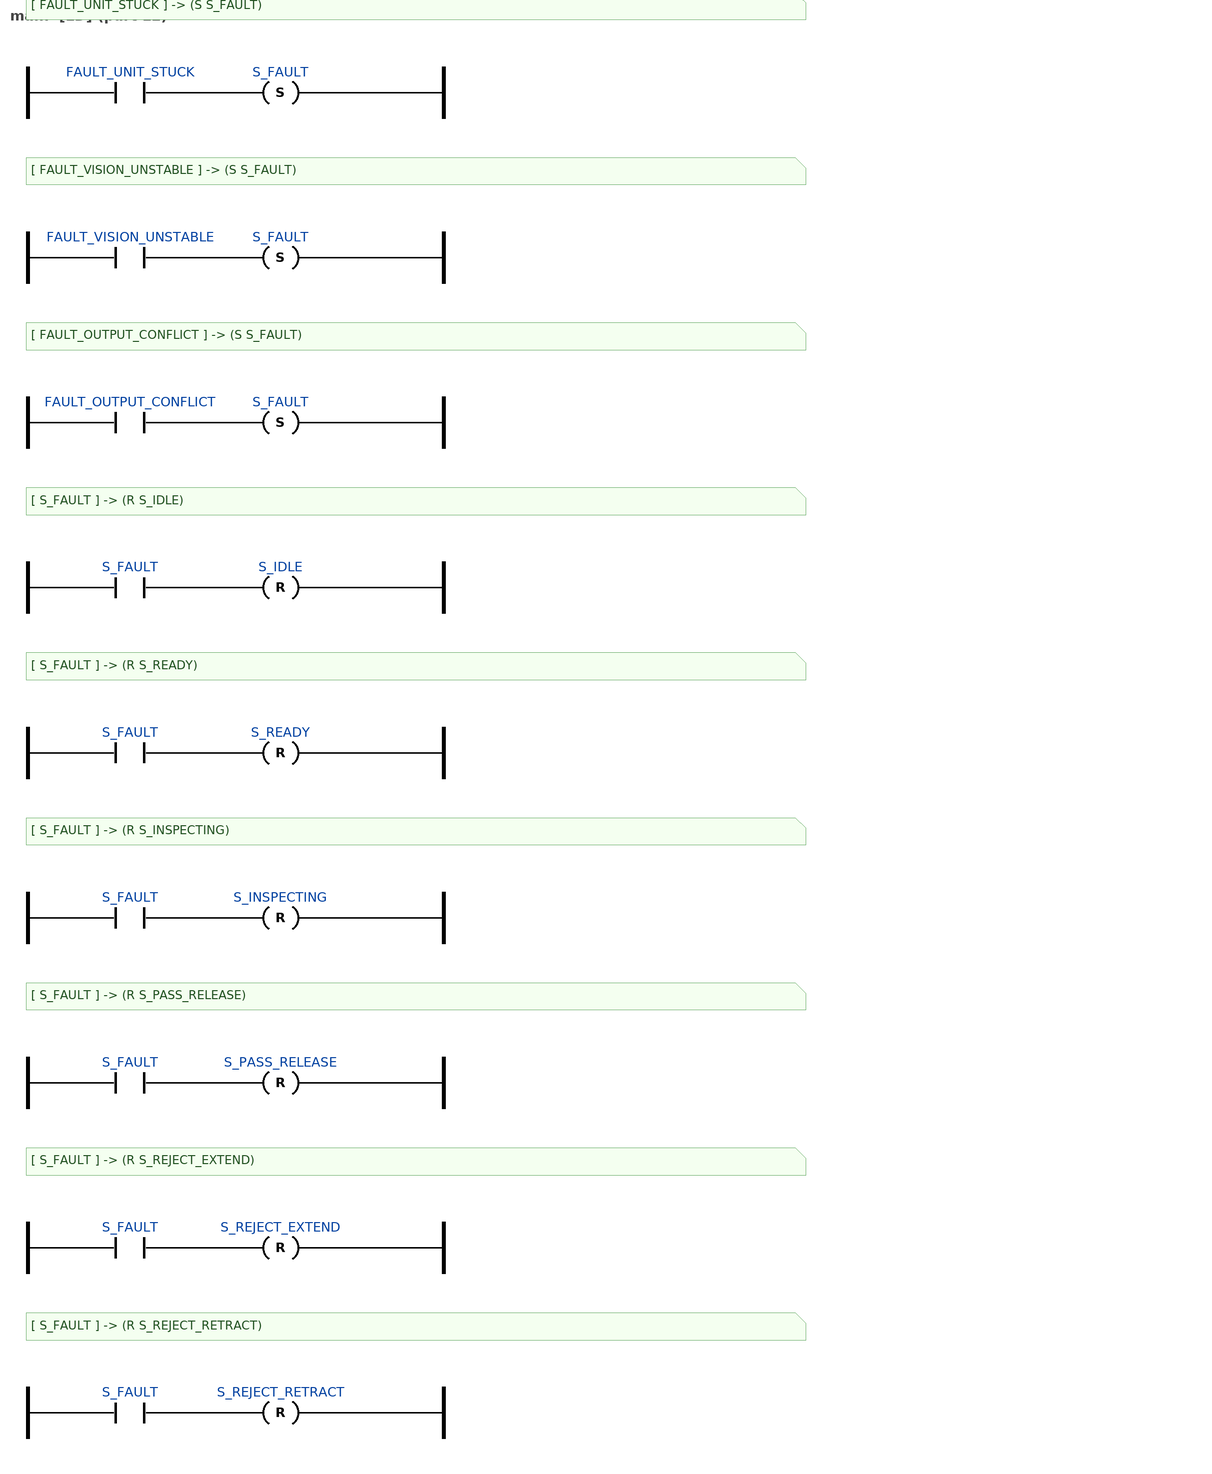
(* [ FAULT_UNIT_STUCK ] -> (S S_FAULT) *)
IF FAULT_UNIT_STUCK THEN S_FAULT := TRUE; END_IF;
(* [ FAULT_VISION_UNSTABLE ] -> (S S_FAULT) *)
IF FAULT_VISION_UNSTABLE THEN S_FAULT := TRUE; END_IF;
(* [ FAULT_OUTPUT_CONFLICT ] -> (S S_FAULT) *)
IF FAULT_OUTPUT_CONFLICT THEN S_FAULT := TRUE; END_IF;
(* [ S_FAULT ] -> (R S_IDLE) *)
IF S_FAULT THEN S_IDLE := FALSE; END_IF;
(* [ S_FAULT ] -> (R S_READY) *)
IF S_FAULT THEN S_READY := FALSE; END_IF;
(* [ S_FAULT ] -> (R S_INSPECTING) *)
IF S_FAULT THEN S_INSPECTING := FALSE; END_IF;
(* [ S_FAULT ] -> (R S_PASS_RELEASE) *)
IF S_FAULT THEN S_PASS_RELEASE := FALSE; END_IF;
(* [ S_FAULT ] -> (R S_REJECT_EXTEND) *)
IF S_FAULT THEN S_REJECT_EXTEND := FALSE; END_IF;
(* [ S_FAULT ] -> (R S_REJECT_RETRACT) *)
IF S_FAULT THEN S_REJECT_RETRACT := FALSE; END_IF;
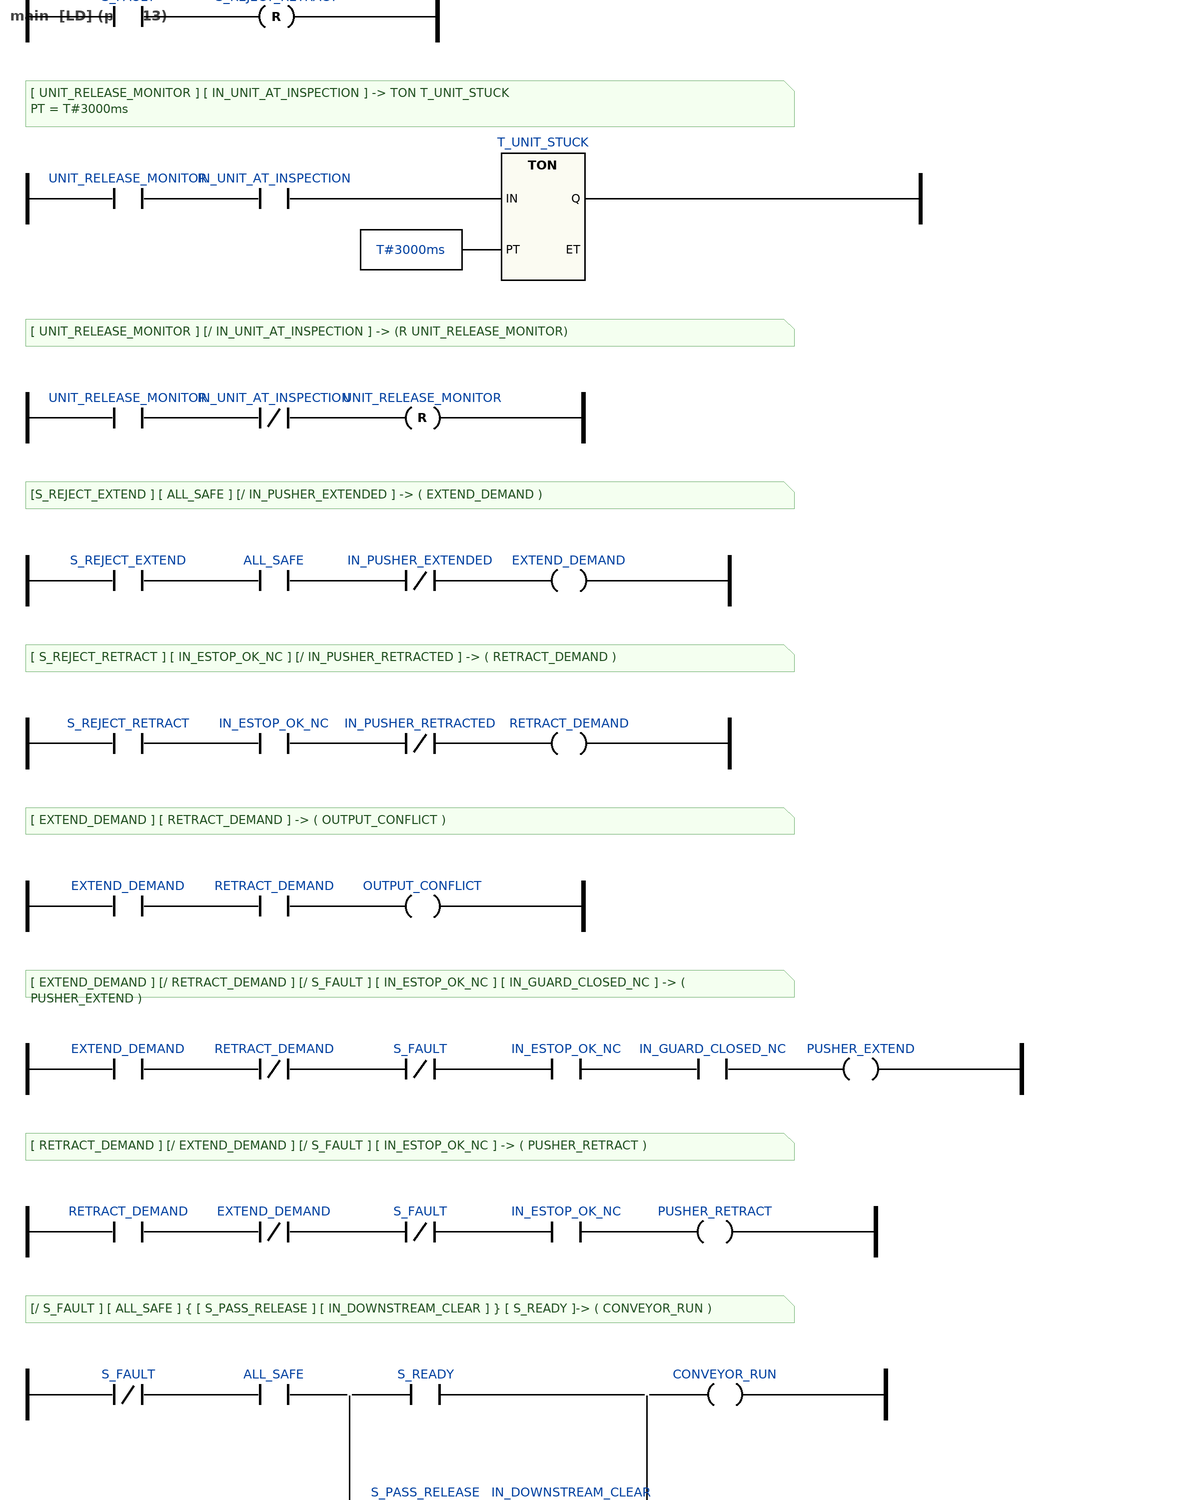
(* [ UNIT_RELEASE_MONITOR ] [ IN_UNIT_AT_INSPECTION ] -> TON T_UNIT_STUCK
PT = T#3000ms *)
(* [ UNIT_RELEASE_MONITOR ] [/ IN_UNIT_AT_INSPECTION ] -> (R UNIT_RELEASE_MONITOR) *)
IF UNIT_RELEASE_MONITOR AND NOT IN_UNIT_AT_INSPECTION THEN UNIT_RELEASE_MONITOR := FALSE; END_IF;
(* [S_REJECT_EXTEND ] [ ALL_SAFE ] [/ IN_PUSHER_EXTENDED ] -> ( EXTEND_DEMAND ) *)
EXTEND_DEMAND := S_REJECT_EXTEND AND ALL_SAFE AND NOT IN_PUSHER_EXTENDED;
(* [ S_REJECT_RETRACT ] [ IN_ESTOP_OK_NC ] [/ IN_PUSHER_RETRACTED ] -> ( RETRACT_DEMAND ) *)
RETRACT_DEMAND := S_REJECT_RETRACT AND IN_ESTOP_OK_NC AND NOT IN_PUSHER_RETRACTED;
(* [ EXTEND_DEMAND ] [ RETRACT_DEMAND ] -> ( OUTPUT_CONFLICT ) *)
OUTPUT_CONFLICT := EXTEND_DEMAND AND RETRACT_DEMAND;
(* [ EXTEND_DEMAND ] [/ RETRACT_DEMAND ] [/ S_FAULT ] [ IN_ESTOP_OK_NC ] [ IN_GUARD_CLOSED_NC ] -> ( PUSHER_EXTEND ) *)
PUSHER_EXTEND := EXTEND_DEMAND AND NOT RETRACT_DEMAND AND NOT S_FAULT AND IN_ESTOP_OK_NC AND IN_GUARD_CLOSED_NC;
(* [ RETRACT_DEMAND ] [/ EXTEND_DEMAND ] [/ S_FAULT ] [ IN_ESTOP_OK_NC ] -> ( PUSHER_RETRACT ) *)
PUSHER_RETRACT := RETRACT_DEMAND AND NOT EXTEND_DEMAND AND NOT S_FAULT AND IN_ESTOP_OK_NC;
(* [/ S_FAULT ] [ ALL_SAFE ] { [ S_PASS_RELEASE ] [ IN_DOWNSTREAM_CLEAR ] } [ S_READY ]-> ( CONVEYOR_RUN ) *)
CONVEYOR_RUN := NOT S_FAULT AND ALL_SAFE AND (S_READY OR S_PASS_RELEASE AND IN_DOWNSTREAM_CLEAR);
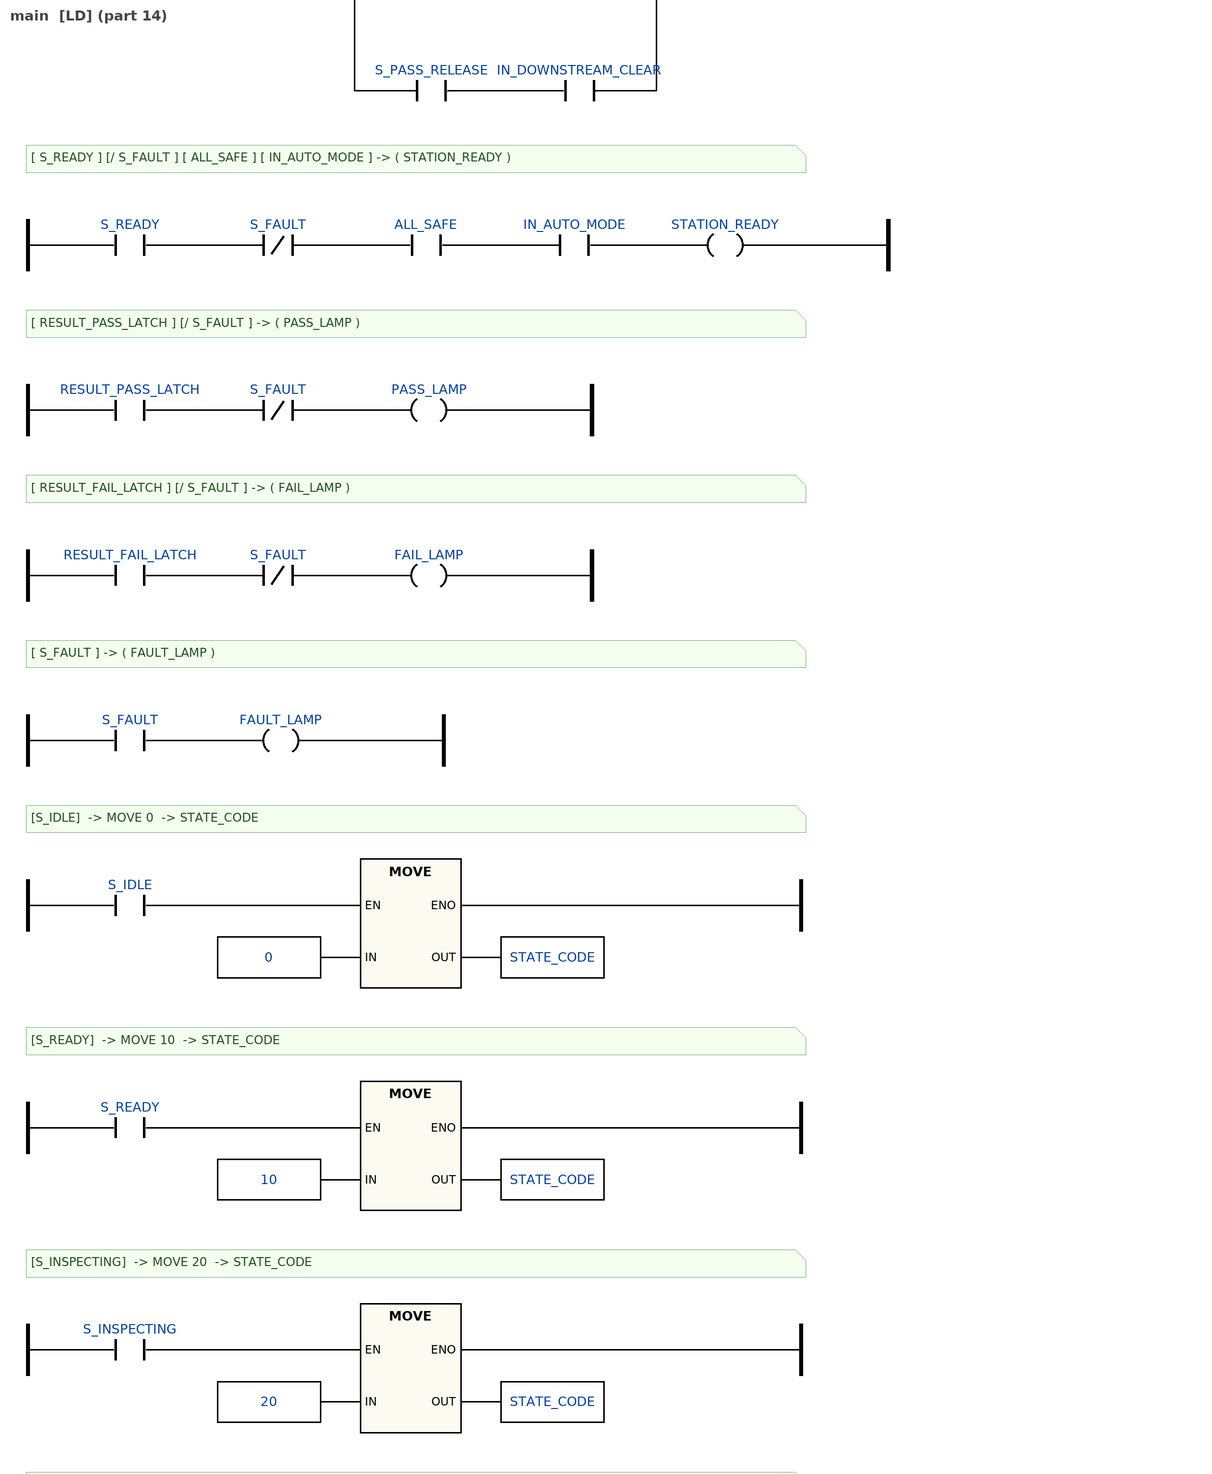
(* [ S_READY ] [/ S_FAULT ] [ ALL_SAFE ] [ IN_AUTO_MODE ] -> ( STATION_READY ) *)
STATION_READY := S_READY AND NOT S_FAULT AND ALL_SAFE AND IN_AUTO_MODE;
(* [ RESULT_PASS_LATCH ] [/ S_FAULT ] -> ( PASS_LAMP ) *)
PASS_LAMP := RESULT_PASS_LATCH AND NOT S_FAULT;
(* [ RESULT_FAIL_LATCH ] [/ S_FAULT ] -> ( FAIL_LAMP ) *)
FAIL_LAMP := RESULT_FAIL_LATCH AND NOT S_FAULT;
(* [ S_FAULT ] -> ( FAULT_LAMP ) *)
FAULT_LAMP := S_FAULT;
(* [S_IDLE]  -> MOVE 0  -> STATE_CODE *)
IF S_IDLE THEN STATE_CODE := 0; END_IF;
(* [S_READY]  -> MOVE 10  -> STATE_CODE *)
IF S_READY THEN STATE_CODE := 10; END_IF;
(* [S_INSPECTING]  -> MOVE 20  -> STATE_CODE *)
IF S_INSPECTING THEN STATE_CODE := 20; END_IF;
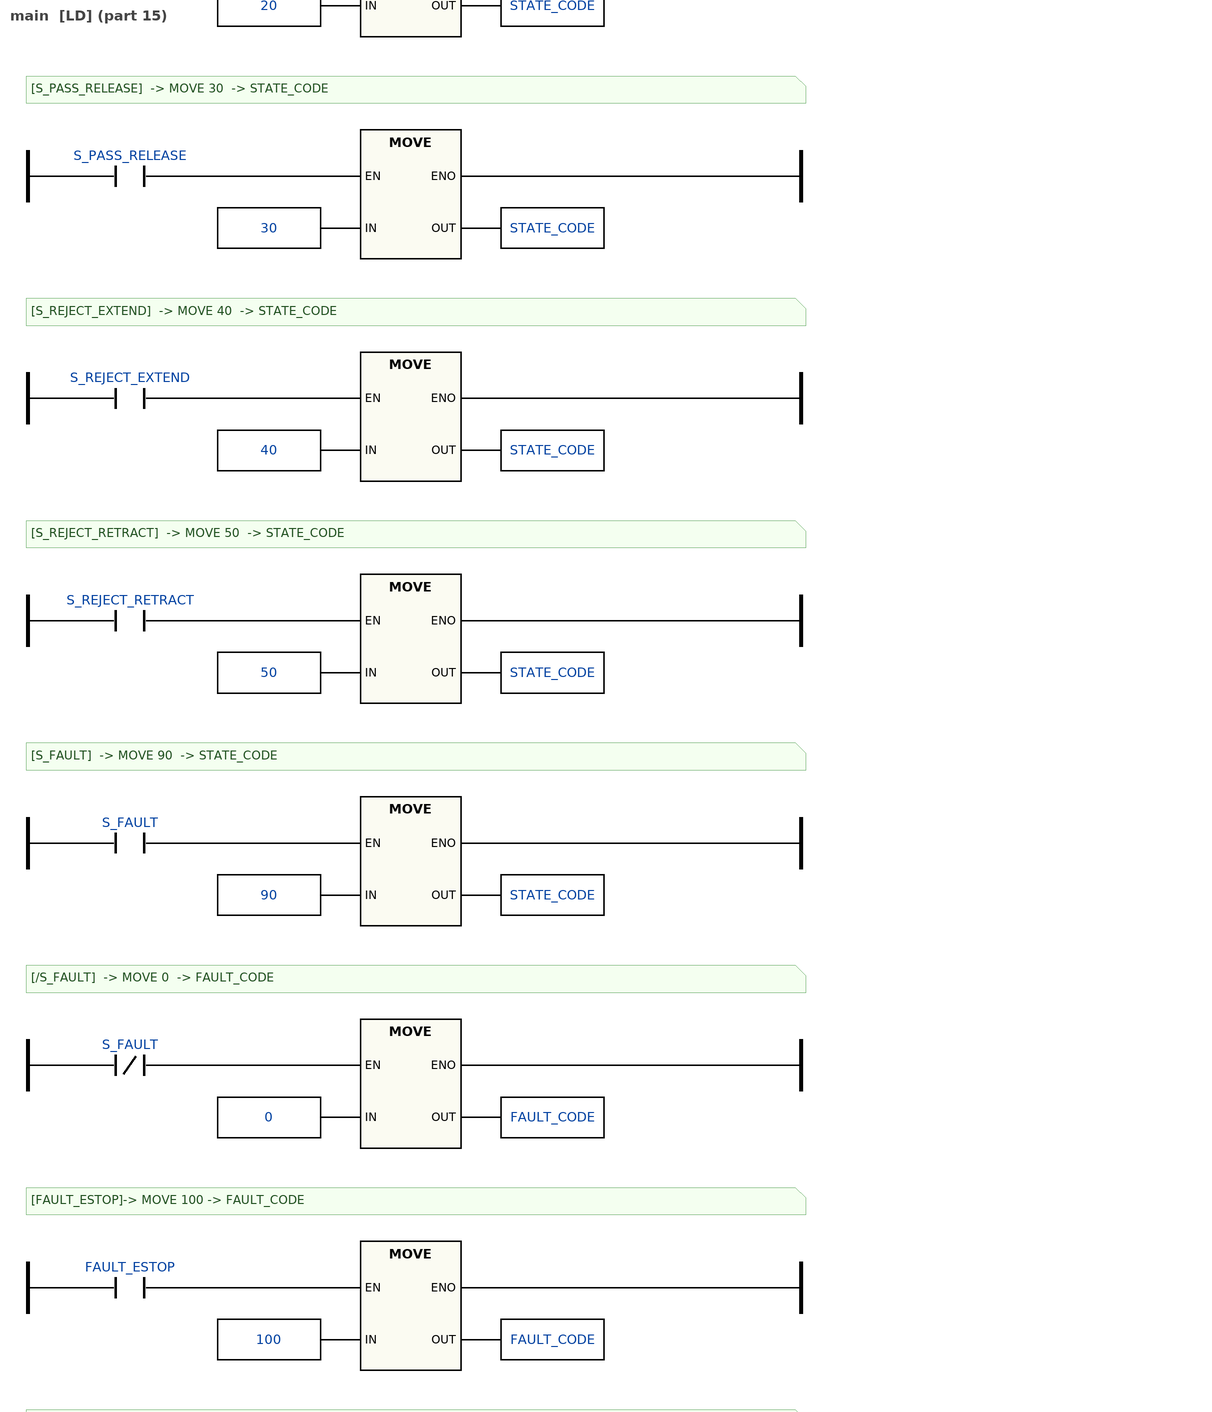
(* [S_PASS_RELEASE]  -> MOVE 30  -> STATE_CODE *)
IF S_PASS_RELEASE THEN STATE_CODE := 30; END_IF;
(* [S_REJECT_EXTEND]  -> MOVE 40  -> STATE_CODE *)
IF S_REJECT_EXTEND THEN STATE_CODE := 40; END_IF;
(* [S_REJECT_RETRACT]  -> MOVE 50  -> STATE_CODE *)
IF S_REJECT_RETRACT THEN STATE_CODE := 50; END_IF;
(* [S_FAULT]  -> MOVE 90  -> STATE_CODE *)
IF S_FAULT THEN STATE_CODE := 90; END_IF;
(* [/S_FAULT]  -> MOVE 0  -> FAULT_CODE *)
IF NOT S_FAULT THEN FAULT_CODE := 0; END_IF;
(* [FAULT_ESTOP]-> MOVE 100 -> FAULT_CODE *)
IF FAULT_ESTOP THEN FAULT_CODE := 100; END_IF;
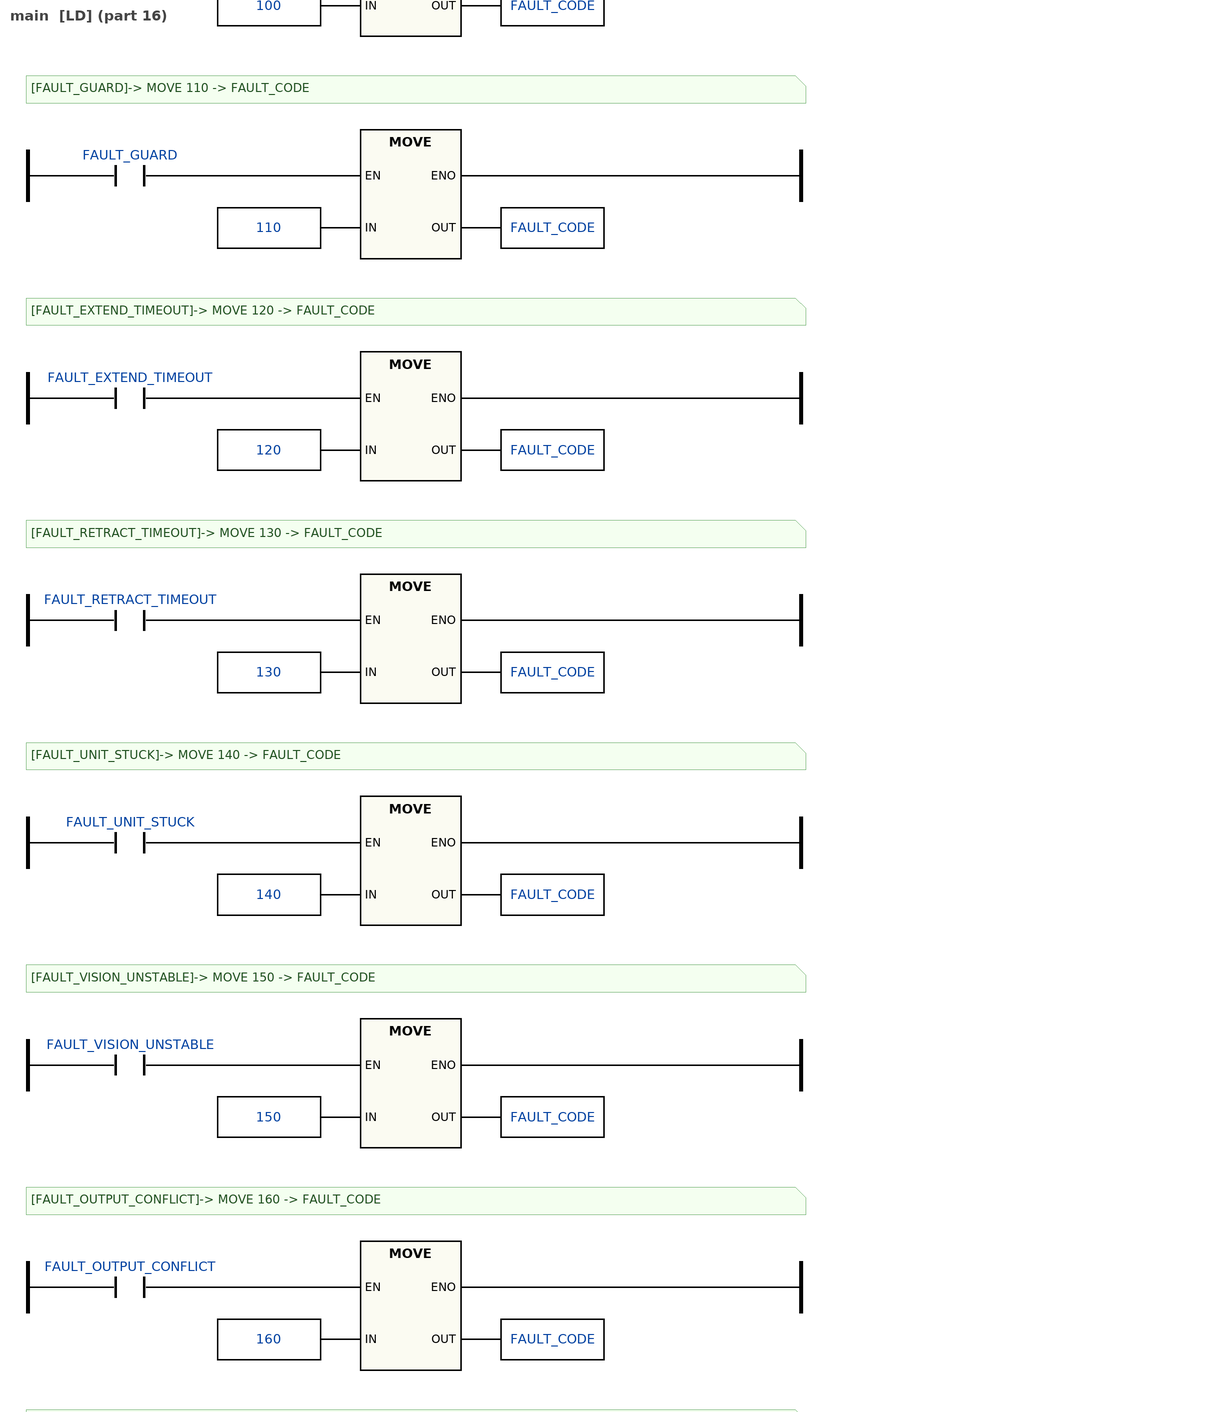
(* [FAULT_GUARD]-> MOVE 110 -> FAULT_CODE *)
IF FAULT_GUARD THEN FAULT_CODE := 110; END_IF;
(* [FAULT_EXTEND_TIMEOUT]-> MOVE 120 -> FAULT_CODE *)
IF FAULT_EXTEND_TIMEOUT THEN FAULT_CODE := 120; END_IF;
(* [FAULT_RETRACT_TIMEOUT]-> MOVE 130 -> FAULT_CODE *)
IF FAULT_RETRACT_TIMEOUT THEN FAULT_CODE := 130; END_IF;
(* [FAULT_UNIT_STUCK]-> MOVE 140 -> FAULT_CODE *)
IF FAULT_UNIT_STUCK THEN FAULT_CODE := 140; END_IF;
(* [FAULT_VISION_UNSTABLE]-> MOVE 150 -> FAULT_CODE *)
IF FAULT_VISION_UNSTABLE THEN FAULT_CODE := 150; END_IF;
(* [FAULT_OUTPUT_CONFLICT]-> MOVE 160 -> FAULT_CODE *)
IF FAULT_OUTPUT_CONFLICT THEN FAULT_CODE := 160; END_IF;
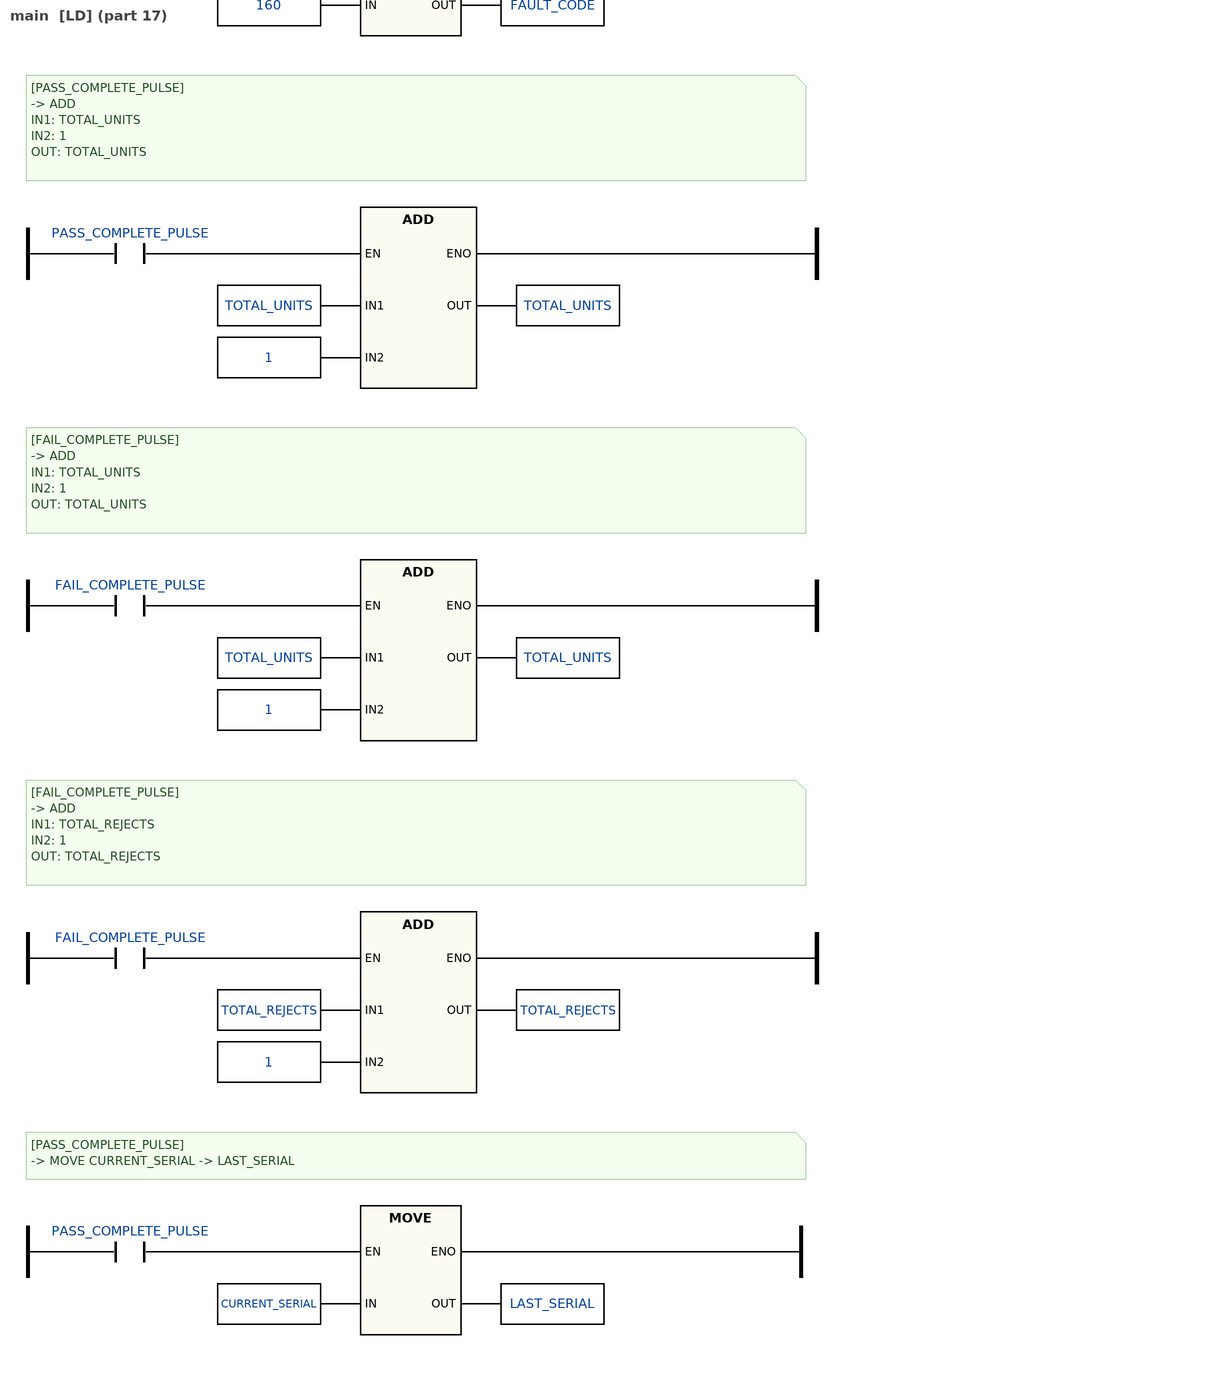
(* [PASS_COMPLETE_PULSE]
    -> ADD
       IN1: TOTAL_UNITS
       IN2: 1
       OUT: TOTAL_UNITS *)
IF PASS_COMPLETE_PULSE THEN TOTAL_UNITS := TOTAL_UNITS + 1; END_IF;
(* [FAIL_COMPLETE_PULSE]
    -> ADD
       IN1: TOTAL_UNITS
       IN2: 1
       OUT: TOTAL_UNITS *)
IF FAIL_COMPLETE_PULSE THEN TOTAL_UNITS := TOTAL_UNITS + 1; END_IF;
(* [FAIL_COMPLETE_PULSE]
    -> ADD
       IN1: TOTAL_REJECTS
       IN2: 1
       OUT: TOTAL_REJECTS *)
IF FAIL_COMPLETE_PULSE THEN TOTAL_REJECTS := TOTAL_REJECTS + 1; END_IF;
(* [PASS_COMPLETE_PULSE]
    -> MOVE CURRENT_SERIAL -> LAST_SERIAL *)
IF PASS_COMPLETE_PULSE THEN LAST_SERIAL := CURRENT_SERIAL; END_IF;
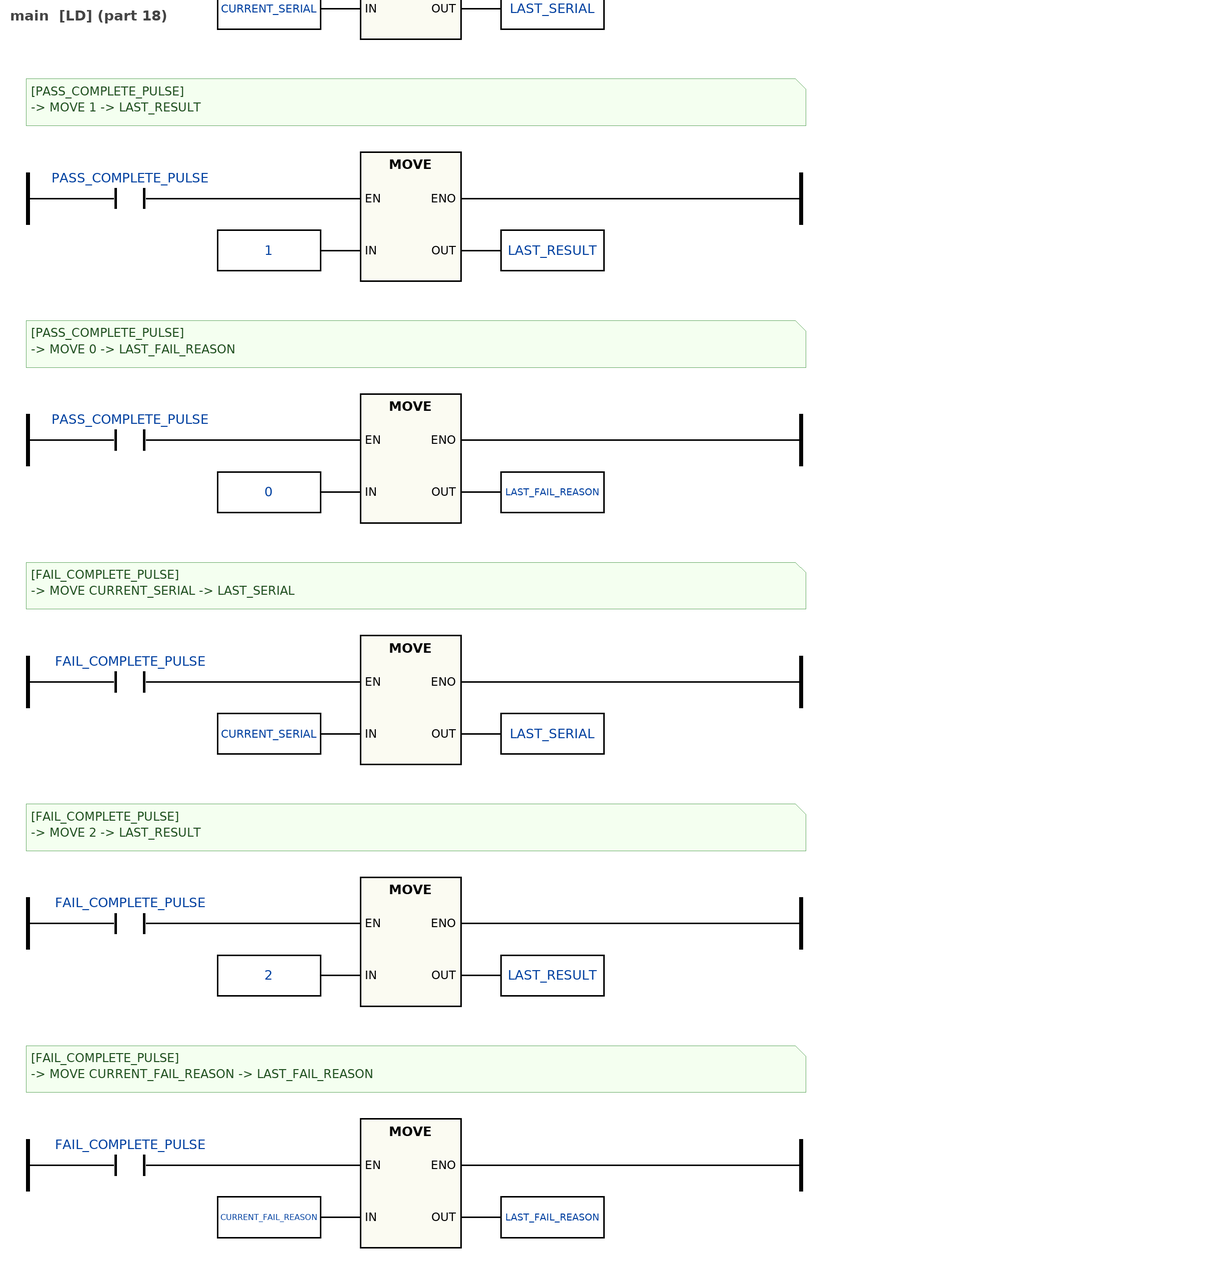
(* [PASS_COMPLETE_PULSE]
    -> MOVE 1 -> LAST_RESULT *)
IF PASS_COMPLETE_PULSE THEN LAST_RESULT := 1; END_IF;
(* [PASS_COMPLETE_PULSE]
    -> MOVE 0 -> LAST_FAIL_REASON *)
IF PASS_COMPLETE_PULSE THEN LAST_FAIL_REASON := 0; END_IF;
(* [FAIL_COMPLETE_PULSE]
    -> MOVE CURRENT_SERIAL -> LAST_SERIAL *)
IF FAIL_COMPLETE_PULSE THEN LAST_SERIAL := CURRENT_SERIAL; END_IF;
(* [FAIL_COMPLETE_PULSE]
    -> MOVE 2 -> LAST_RESULT *)
IF FAIL_COMPLETE_PULSE THEN LAST_RESULT := 2; END_IF;
(* [FAIL_COMPLETE_PULSE]
    -> MOVE CURRENT_FAIL_REASON -> LAST_FAIL_REASON *)
IF FAIL_COMPLETE_PULSE THEN LAST_FAIL_REASON := CURRENT_FAIL_REASON; END_IF;
T_VISION_STABLE(IN := S_INSPECTING AND IN_VISION_RESULT_VALID AND NOT VISION_CHANGED, PT := T#250ms);
T_VISION_UNSTABLE(IN := S_INSPECTING AND IN_VISION_RESULT_VALID AND VISION_UNSTABLE_LATCH, PT := T#1000ms);
T_PASS_RELEASE(IN := S_PASS_RELEASE, PT := T#500ms);
T_EXTEND_TIMEOUT(IN := S_REJECT_EXTEND AND NOT IN_PUSHER_EXTENDED, PT := T#1500ms);
T_REJECT_SETTLE(IN := S_REJECT_EXTEND AND IN_PUSHER_EXTENDED, PT := T#250ms);
T_RETRACT_TIMEOUT(IN := S_REJECT_RETRACT AND NOT IN_PUSHER_RETRACTED, PT := T#1500ms);
T_UNIT_STUCK(IN := UNIT_RELEASE_MONITOR AND IN_UNIT_AT_INSPECTION, PT := T#3000ms);
END_PROGRAM
